// ---- POUs/Tc2 Objects/Signals/Watchdog/FB_SignalWatchdog.TcPOU
FUNCTION_BLOCK FB_SignalWatchdog
VAR_INPUT
	(* Input variables / Eingang Variablen *)
	bEnable					:BOOL;						(* Enable FB signal *)
	bIn						:BOOL;						(* Input signal *)
	tWatchdog				:TIME := t#0s;					(* Watchdog time *)
END_VAR
VAR_OUTPUT
	(* Output variables / Ausgang Variablen *)
	bOut					:BOOL;						(* Output signal *)
	bAlarm					:BOOL;						(* Alarm signal *)
END_VAR
VAR
	(* Enummerations *)

	(* Variables *)


	(* References *)

	(* Interfaces *)

	(* Instances *)
	tofWatchdog				:TOF;

END_VAR

IF NOT bEnable
THEN
	bOut := FALSE;
	bAlarm := FALSE;                       (* Alarm active *)
	
	tofWatchdog(
		IN := tofWatchdog.ET > t#0ms,
	         PT := t#0ms
	);
	
	tofWatchdog(IN := FALSE,
	             PT := t#0ms);

	RETURN;
END_IF;

tofWatchdog(					 (* Dealy input signal *)
	IN := bIn,
	PT := tWatchdog
);

bOut := tofWatchdog.Q;

bAlarm := NOT tofWatchdog.Q;                       (* Set alarm *)

END_FUNCTION_BLOCK

// ---- POUs/Machine/Group_0000 - General/Gr00Control/Gr00Signals/FB_Gr00Signals.TcPOU
FUNCTION_BLOCK FB_Gr00Signals
(*

The function block used to control general signals of the machine.

Constructor: 		Patryk Panylo
Company:		E. Riexinger GmbH
Date:			28.04.2015
Version:			1.00

Date:			Revision:		Who:				Comment
dd.mm.yyyy		x.xx			Initials			comment

*)
VAR_INPUT
	(* Input variables / Eingang Variablen *)
	etMachineMode				:ET_MachineMode;			(* Machine mode *)
	etMachineState				:ET_MachineState;			(* Machine state *)
	bMachineRunning				:BOOL;						(* Machine running / Maschine lauft *)
	stAlarm						:ST_Alarm;					(* Current status of alarms *)
END_VAR
VAR_OUTPUT
	(* Output variables / Ausgang Variablen *)
	bBulbRed					:BOOL;						(* Signal column bulb "stop" or "error" / Signallampe "Stop" oder "Fehler" *)
	bBulbYellow					:BOOL;						(* Signal column bulb "warning" or "message" / Signallampe "Warnung" oder "Message" *)
	bBulbGreen					:BOOL;						(* Signal column bulb "automatic" / Signallampe "Automatik" *)
	bBulbBtnStop					:BOOL;						(* Signal button bulb "stop" / Signallampe "Stop" *)
	bBulbBtnHome				:BOOL;						(* Signal button bulb "home" / Signallampe "Grundstellung" *)
	bBulbBtnStart					:BOOL;						(* Signal button bulb "start" / Signallampe "Start" *)
	bHorn						:BOOL;						(* Signal horn / Signalhupe *)
	stBlinker						:ST_Blinker;
END_VAR
VAR_IN_OUT
	(* Input Output variables / Ausgang Variablen *)

END_VAR
VAR
	(* Enummerations *)

	(* Variables *)
	nIdxHorn						:INT;

	(* References *)

	(* Interfaces *)

	(* Instances *)
	fbBlinker						:FB_Blinker;
	rtHorn						:R_TRIG;
	tonDelay						:TON;

END_VAR
VAR CONSTANT
	nHornRepeat					:INT := 3;
END_VAR


A_Blinker();
A_SignalColumn();
A_SignalButton();
A_Horn();

ACTION A_Blinker:

(* Blinker frequency division *)
fbBlinker(
    stBlinker => stBlinker
);
END_ACTION

ACTION A_Horn:

(* Signal horn / Signalhupe *)
IF stBlinker.Q1
     AND nIdxHorn < nHornRepeat
THEN
	bHorn := (stAlarm.bFatalError OR stAlarm.bError);

ELSIF NOT stBlinker.Q1
THEN
	bHorn := FALSE;
END_IF;

rtHorn(CLK := bHorn);
IF rtHorn.Q
THEN
	nIdxHorn := nIdxHorn + 1;
END_IF;

tonDelay(
	IN := nIdxHorn >= nHornRepeat,
	PT := t#60s
);

IF (tonDelay.Q
    AND nHornRepeat > 0)
    OR NOT (stAlarm.bFatalError OR stAlarm.bError)
THEN
	nIdxHorn := 0;
END_IF;
END_ACTION

ACTION A_SignalButton:

(* Signal button bulb "stop" / Signallampe "Stop" *)
bBulbBtnStop := bBulbRed;

(* Signal button bulb "home" / Signallampe "Grundstellung" *)
bBulbBtnHome := (
	(etMachineMode = ET_MachineMode_eHome
	 AND NOT bMachineRunning)
	OR
	(etMachineMode = ET_MachineMode_eHome
	 AND bMachineRunning
	 AND stBlinker.Q1)
);

(* Signal button bulb "start" / Signallampe "Start" *)
bBulbBtnStart := (
	(etMachineMode = ET_MachineMode_eAutomatic
	 AND bMachineRunning)
	OR
	(etMachineMode = ET_MachineMode_eHome
	 AND bMachineRunning
	 AND NOT stBlinker.Q1)
);
END_ACTION

ACTION A_SignalColumn:

(* Signal column bulb "stop" or "error" / Signallampe "Stop" oder "Fehler" *)
bBulbRed := SEL(
	stAlarm.bFatalError OR stAlarm.bError,
	NOT bMachineRunning,
	stBlinker.Q1
);

(* Signal column bulb "warning" or "message" / Signallampe "Warnung" oder "Message" *)
bBulbYellow := (
	NOT stBlinker.Q1
	AND (stAlarm.bWarning OR stAlarm.bMessage)
);

(* Signal column bulb "automatic" / Signallampe "Automatik" *)
bBulbGreen := (
	(etMachineMode = ET_MachineMode_eAutomatic
	 AND bMachineRunning)
	OR
	(etMachineMode = ET_MachineMode_eHome
	 AND bMachineRunning
	 AND stBlinker.Q1)
);
END_ACTION

END_FUNCTION_BLOCK

// ---- POUs/Tc2 Objects/Signals/Generators/FB_Blinker.TcPOU
FUNCTION_BLOCK FB_Blinker
(*

Frequency division

Constructor: 		Patryk Panylo
Company:		E. Riexinger GmbH
Date:			14.11.2012
Version:			1.00

Date:			Revision:		Who:				Comment
dd.mm.yyyy		x.xx			Initials			comment

*)

VAR_INPUT
	tPeriod				:TIME := T#250MS;				(* Blink period *)
	bReset				:BOOL;						(* Reset *)
END_VAR
VAR_OUTPUT
	stBlinker				:ST_Blinker;
END_VAR
VAR
	byInc				:BYTE;
	rtTriger				:R_TRIG;
	ton1					:TON;
	ton2					:TON;
END_VAR

IF bReset
THEN
	byInc := 0;

	ton1(IN := FALSE);
	ton2(IN := FALSE);

	stBlinker.Q0 := 0;
	stBlinker.Q1 := 0;
	stBlinker.Q2 := 0;
	stBlinker.Q3 := 0;
	stBlinker.Q4 := 0;
	stBlinker.Q5 := 0;
	stBlinker.Q6 := 0;
	stBlinker.Q7 := 0;
	
	RETURN;	
END_IF

ton1(IN := NOT ton2.Q, PT:= tPeriod/2);
ton2(IN := ton1.Q, PT := tPeriod/2);

rtTriger(CLK := ton1.Q);
IF rtTriger.Q THEN
	byInc := byInc + 1;
END_IF;

stBlinker.Q0 := byInc.0;
stBlinker.Q1 := byInc.1;
stBlinker.Q2 := byInc.2;
stBlinker.Q3 := byInc.3;
stBlinker.Q4 := byInc.4;
stBlinker.Q5 := byInc.5;
stBlinker.Q6 := byInc.6;
stBlinker.Q7 := byInc.7;

END_FUNCTION_BLOCK

// ---- POUs/Machine/Group_0000 - General/Gr00Control/Gr00Utility/FB_Gr00Utility.TcPOU
FUNCTION_BLOCK FB_Gr00Utility
(*

The function block used to control general utility of the machine.

Constructor: 		Patryk Panylo
Company:		E. Riexinger GmbH
Date:			28.04.2015
Version:			1.00

Date:			Revision:		Who:				Comment
dd.mm.yyyy		x.xx			Initials			comment

*)
VAR_INPUT
	(* Input variables / Eingang Variablen *)
	bSignalStart					:BOOL;						(* Signal "Start" / Signal "Start" *)
	bSignalStop					:BOOL;						(* Signal "Stop" / Signal "Stop" *)
	bSignalAbort					:BOOL;						(* Signal "Abort" / Signal "Abort" *)
	bSignalHome					:BOOL;						(* Signal "Home" / Signal "Grundstellung" *)
	bSignalReference				:BOOL;						(* Signal "Reference" / Signal "Referenz" *)
	bSignalReset					:BOOL;						(* Signal "Reset" / Signal "Reset *)
	bSignalMachinePurge			:BOOL;						(* Machine purge *)
	bAutoStartRelease			:BOOL;						(* Auto start release *)
	bHomeStartRelease			:BOOL;						(* Home start release *)
	bAutoToHome				:BOOL;						(* If auto completed go to home *)
	bHomeCompleted				:BOOL;						(* Home completed signal *)
	bAutoCompleted				:BOOL;						(* Auto completed signal *)
	bAllDoorsClosed 				:BOOL;						(* All doors closed *)
	bAllDoorsLocked 				:BOOL;						(* All doors locked *)
	bLightCurtainOk				:BOOL;						(* Light curtain ok *)
	bExeCounter					:BOOL;						(* Execute counter *)
	bResetCounterUser			:BOOL;						(* Reset counter user *)
	bStartTime					:BOOL;						(* Start measurement of cylce time *)
	bStopTime					:BOOL;						(* Stop measurement of cylce time *)
	bLifetimeOn					:BOOL;						(* Lifetime on *)
	bResetLifetimeAll				:BOOL; 						(* Reset all counters *)
	sLifetimeFilePath				:STRING;					(* File path for life time *)
	sLifetimeFileName			:STRING;					(* File name for life time *)
	bWritePersistent				:BOOL;						(* Write persistent data *)
	bDownTraceDataExe 			:BOOL;						(* Download traceability data *)
	stTraceability					:ST_Traceability;				(* Traceability data *)
	tAdsTimeOut 					:TIME := t#2s;					(* Timout for ads commands *)
END_VAR
VAR_OUTPUT
	(* Output variables / Ausgang Variablen *)
	etMachineMode				:ET_MachineMode;			(* Machine mode *)
	etMachineState				:ET_MachineState;			(* Machine state *)
	bModeAutomatic				:BOOL;						(* Machine mode automatic *)
	bModeHome					:BOOL;						(* Machine mode home *)
	bModeManual				:BOOL;						(* Machine mode manual *)
	bMachineRunning				:BOOL;						(* Machine running *)
	bMachineStandstill			:BOOL;						(* Machine standstill *)
	bMachinePurge				:BOOL;						(* Machine purge *)
	bConfirmAlarm				:BOOL;						(* Alarm confirm *)
	rActOverride					:REAL;						(* Actual override *)
	lrLifetimeAll					:LREAL;						(* Lifetime *)
	lrLifetimeAfterTrunOn			:LREAL;						(* Time after turn on *)
	lrActCycleTime				:LREAL;						(* Actual cycle time *)
	dwCycleTime					:DWORD;					(* Cycletime in 0.01sec / Zykluszeit in 0.01Sekunden *)
END_VAR
VAR_IN_OUT
	(* Input Output variables / Ausgang Variablen *)
	etMachineModeReq			:ET_MachineMode;			(* Machine mode request *)
	rGlobalOverride				:REAL;						(* Global override *)
	udnCounterTotal				:UDINT;						(* Total counter *)
	udnCounterUser				:UDINT;						(* Total counter *)
END_VAR
VAR
	(* Enummerations *)

	(* Variables *)
	nIRHSCtrlCnt					:INT;
	nIRHSZoneCnt				:INT;
	lrIRHSSetpointLeftSide			:LREAL;
	lrIRHSSetpointRightSide		:LREAL;

	bTraceExe					:BOOL;
	ftTraceExe					:F_TRIG;
	rtDownTraceDataExe			:R_TRIG;
	rtDownTraceDataReset		:R_TRIG;
	udnTraceSampleCnt			:UDINT;
	udnTraceDataCnt				:UDINT;

	(* References *)

	(* Interfaces *)

	(* Instances *)
	fbModeSelector				:FB_ModeSelector;			(* Mode selector *)
	fbOverride					:FB_Override;					(* Override *)
	fbLifetime					:FB_TimeHoursCounter;		(* Machine lifetime *)
	fbCounterTotal				:FB_Counter;					(* Counter total *)
	fbCounterUser				:FB_Counter;					(* Counter user *)
	rtResetCounterUser			:R_TRIG;						(* Reset counter user *)
	fbCylceTime					:FB_Timer;					(* Machine cycle time *)
	fbSUPS						:FB_S_UPS_CX51x0;			(*  The function block FB_S_UPS_CX51x0 can be used on CX devices with one-second UPS to control the one-second UPS from the PLC *)
	fbWritePersistentData			:WritePersistentData;			(*  Write Persistent *)
	fbGetCurTaskIdx				:GETCURTASKINDEX;			(* This function block finds the task index of the task from which it is called *)
	fbRTC						:FB_RTC;					(* Get current time *)
	fbTraceability					:FB_Traceability;				(* Traceability *)
	rtMachinePurge				:R_TRIG;
	SystemTaskInfoArr: INT;
END_VAR


A_OperationMode();
A_Override();
A_Counter();
A_CycleTime();
A_MachinePurge();
A_Persistent();
A_PlcTaskSystemInfo();
A_RTC();
A_Traceability();

ACTION A_Counter:

(* Hours counter *)
fbLifetime(
	bEnable := TRUE,
	bDeleteAll := bResetLifetimeAll,
	sAmsNetId := sgAmsNetId,
	bCount := bLifetimeOn,
	bSave := FALSE,
	sFilePath := sLifetimeFilePath,
	sFileName := sLifetimeFileName,
	tSaveIntervall := t#5m,
	tTimeout := tAdsTimeOut,
	lrAllOverHours => lrLifetimeAll,
	lrNoRetainHours => lrLifetimeAfterTrunOn,
 );

(* General counter *)
fbCounterTotal(
	bEnable := TRUE,
	bExecute := bExeCounter,
	bReset := fbCounterTotal.bOverflow,
	udnCounter := udnCounterTotal
);

rtResetCounterUser(CLK:= bResetCounterUser);

fbCounterUser(
	bEnable := TRUE,
	bExecute := bExeCounter,
	bReset := rtResetCounterUser.Q
			 OR fbCounterUser.bOverflow,
	udnCounter := udnCounterUser
);
END_ACTION

ACTION A_CycleTime:

(* Cylce time *)
fbCylceTime(
	bEnable := TRUE,
	bReset := FALSE,
	bStartStop := bStartTime
			        AND bModeAutomatic,
	bStop := bStopTime
		        OR bMachineStandstill,
	tMaxTime := ,
	stRefTime => ,
	stActTime => ,
	stRestTime =>
);

dwCycleTime := fbCylceTime.stActTime.dwDeciSec;
END_ACTION

ACTION A_MachinePurge:

rtMachinePurge(CLK := 	bSignalMachinePurge);

IF NOT bModeAutomatic
     OR bAutoCompleted
THEN
	bMachinePurge := FALSE;

ELSIF rtMachinePurge.Q
THEN
	bMachinePurge := TRUE;
END_IF
END_ACTION

ACTION A_OperationMode:

(* Operation mode control *)
fbModeSelector(
	bStart := bSignalStart,
	bStop := bSignalStop,
	bAbort := bSignalAbort,
	bHome := bSignalHome,
	bReset := bSignalReset,
	bReference := bSignalReference,
	bAutoStartRelease := bAutoStartRelease,
	bHomeStartRelease := bHomeStartRelease,
	bAutoToHome := bAutoToHome,
	bHomeCompleted := bHomeCompleted,
	bAutoCompleted := bAutoCompleted,
	bAllDoorsClosed  := bAllDoorsClosed,
	bAllDoorsLocked := bAllDoorsLocked,
	bLightCurtainOk := bLightCurtainOk,
	etMachineMode => etMachineMode,
	etMachineState => etMachineState,
	bModeAutomatic => bModeAutomatic,
	bModeHome => bModeHome,
	bModeManual => bModeManual,
	bMachineRunning => bMachineRunning,
	bMachineStandstill => bMachineStandstill,
	bConfirmAlarm => bConfirmAlarm,
	etMachineModeReq := etMachineModeReq
);
END_ACTION

ACTION A_Override:

(* Override control *)
fbOverride(
	bEnable := TRUE,
	bBypassAccDec := bModeManual,
	bSetOverideMax := bModeAutomatic,
	rAcc := rgGr00AdsOverrideAcc,
	rDec := rgGr01AdsOverrideDec,
	rSetOverride := rGlobalOverride,
	rActOverride => rActOverride
);
END_ACTION

ACTION A_Persistent:

(*  The function block FB_S_UPS_CX51x0 can be used on CX devices with one-second UPS to control the one-second UPS from the PLC *)
fbSUPS(
	sNetID := sgAmsNetId,													(* AmsNetID of the controller. *)
	iPLCPort := AMSPORT_R0_PLC_RTS1,									(* Port number of the PLC runtime system (AMSPORT_R0_PLC_RTS1 = 801, AMSPORT_R0_PLC_RTS2 = 811, AMSPORT_R0_PLC_RTS3 = 821, AMSPORT_R0_PLC_RTS4 = 831). *)
	iUPSPort := 16#588,													(* Port number via which the UPS status is read (standard value is 16#588) *)
	tTimeout := DEFAULT_ADS_TIMEOUT,									(* ADS Timeout *)
	eUpsMode := eSUPS_WrPersistData_Shutdown,							(* The eUpsMode defines whether persistent data are to be written and whether a QuickShutdown is to be performed.
																		Standard value is eSUPS_WrPersistData_Shutdown, i.e. with writing of the persistent data and then QuickShutdown. See E_S_UPS_Mode. *)
	ePersistentMode := SPDM_2PASS,										(* Mode for the writing of the persistent data. Standard value is SPDM_2PASS *)
	tRecoverTime := t#10s													(* Time after which the UPS reverts to the PowerOK status in the case of UPS modes without shutdown.
																	   	    The tRecoverTime must be somewhat longer than the maximum holding time of the UPS, since the UPS switches off even when the voltage returns. *)
);


(* If persistent variables are defined in one of the PLC's runtime systems, then their current values are stored in a file in the TwinCAT\Boot directory when the TwinCAT system stops (after the last PLC cycle). *)
fbWritePersistentData(
	NETID := sgAmsNetId,
	PORT := AMSPORT_R0_PLC_RTS1,
	START := bWritePersistent
			   AND NOT fbWritePersistentData.BUSY,
	TMOUT := DEFAULT_ADS_TIMEOUT
);
END_ACTION

ACTION A_PlcTaskSystemInfo:

fbGetCurTaskIdx();

// lrActCycleTime := UDINT_TO_LREAL(SystemTaskInfoArr[fbGetCurTaskIdx.index].cycleTime) / 10000000;




fbGetCurTaskIdx();

GVL._PlcTaskSystemInfo := _TaskInfo[fbGetCurTaskIdx.index];

lrActCycleTime := UDINT_TO_LREAL(_TaskInfo[fbGetCurTaskIdx.index].CycleTime) / 10000000;
END_ACTION

ACTION A_RTC:

fbRTC(
	stDateTime => stgGr00DateTime
);
END_ACTION

ACTION A_Traceability:

stTraceability.sDateTime := stgGr00DateTime.sDateTime;

stTraceability.stSettings.sPath := sTracePath(*CONCAT(CONCAT(sTracePath,fbRTC.sDate),'\')*);
stTraceability.stSettings.sFileName := stgGr00DateTime.sDateTime;
stTraceability.stSettings.sFileExtension := sTraceFileExtension;

rtDownTraceDataReset(
	CLK := bModeAutomatic
);

IF rtDownTraceDataReset.Q
THEN
	udnTraceSampleCnt := 0;
	MEMSET(ADR(stTraceability.arstData), 0, SIZEOF(stTraceability.arstData));
END_IF

rtDownTraceDataExe(
	CLK := bTraceEnable
		    AND bDownTraceDataExe
);

IF rtDownTraceDataExe.Q
     AND udnTraceSampleCnt < udnTraceSampleMax
THEN
	udnTraceDataCnt := 0;
	udnTraceSampleCnt := udnTraceSampleCnt +1;
	(*1*)
	udnTraceDataCnt := udnTraceDataCnt + 1;
	stTraceability.arstData[udnTraceSampleCnt,udnTraceDataCnt].sName := 'Time';
	stTraceability.arstData[udnTraceSampleCnt,udnTraceDataCnt].sValue := stgGr00DateTime.sDateTime;
	stTraceability.arstData[udnTraceSampleCnt,udnTraceDataCnt].sUnit := '';

	(*2*)
	udnTraceDataCnt := udnTraceDataCnt + 1;
	stTraceability.arstData[udnTraceSampleCnt,udnTraceDataCnt].sName := 'Cntr';
	stTraceability.arstData[udnTraceSampleCnt,udnTraceDataCnt].sValue := UDINT_TO_STRING(stgGr00HMI.stPLCTOHMI.udnCounterTotal);
	stTraceability.arstData[udnTraceSampleCnt,udnTraceDataCnt].sUnit := '';

END_IF

(*ftTraceExe(CLK := bgGr00ModeAutomatic);*)
fbTraceability(
	bEnable := bTraceEnable,
	bExecute := bAutoCompleted
			     (*OR
			     (NOT bAutoCompleted
			      AND (bSignalStop OR bSignalAbort)
			      AND ftTraceExe.Q)*)
			     OR bTraceExe,
	stTraceability := stTraceability
);
END_ACTION

END_FUNCTION_BLOCK

// ---- POUs/Tc2 Objects/Automation/OperationMode/FB_ModeSelector.TcPOU
FUNCTION_BLOCK FB_ModeSelector
(*

The function block used to control opration mode.

Constructor: 		Patryk Panylo
Company:		E. Riexinger GmbH
Date:			23.04.2015
Version:			1.00

Date:			Revision:		Who:				Comment
dd.mm.yyyy		x.xx			Initials			comment

*)
VAR_INPUT
	(* Input variables / Eingang Variablen *)
	bStart					:BOOL;						(* Signal start *)
	bStop					:BOOL;						(* Signal stop *)
	bAbort					:BOOL;						(* Signal abort *)
	bHome					:BOOL;						(* Signal home *)
	bReference				:BOOL;						(* Signal reference *)
	bReset					:BOOL;						(* Signal reset *)
	bAutoStartRelease		:BOOL;						(* Auto start release *)
	bHomeStartRelease		:BOOL;						(* Home start release *)
	bAutoToHome			:BOOL;						(* If auto completed go to home *)
	bHomeCompleted			:BOOL;						(* Home completed *)
	bAutoCompleted			:BOOL;						(* Auto completed *)
	bAllDoorsClosed 			:BOOL;						(* All doors closed *)
	bAllDoorsLocked 			:BOOL;						(* All doors locked *)
	bLightCurtainOk			:BOOL;						(* Light curtain ok *)
END_VAR
VAR_OUTPUT
	(* Output variables / Ausgang Variablen *)
	etMachineMode			:ET_MachineMode;			(* Machine mode enum variable *)
	etMachineState			:ET_MachineState;			(* Machine state enum variable *)
	bModeAutomatic			:BOOL;						(* Machine mode automatic *)
	bModeHome				:BOOL;						(* Machine mode home *)
	bModeManual			:BOOL;						(* Machine mode manual *)
	bMachineRunning			:BOOL;						(* Machine running *)
	bMachineStandstill		:BOOL;						(* Machine standstill *)
	bConfirmAlarm			:BOOL;						(* Confirm alarm *)
END_VAR
VAR_IN_OUT
	etMachineModeReq		:ET_MachineMode;			(* Machine mode request enum variable *)
END_VAR
VAR
	(* Enummerations *)

	(* Variables *)
	etMachinePrvState		:ET_MachineState;			(* Machine previous active state enum variable *)
	bModeExecute			:BOOL;						(* Mode execute *)
	bSafetyCompleted		:BOOL;						(* Safety completed *)

	(* References *)

	(* Interfaces *)

	(* Instances *)
	rtStart					:R_TRIG;
	rtStop					:R_TRIG;
	rtAbort					:R_TRIG;
END_VAR


bConfirmAlarm := bReset;
bSafetyCompleted := bAllDoorsLocked				(* Safety completed *)
				      AND bLightCurtainOk;

IF bHome
THEN
	etMachineModeReq := ET_MachineMode_eHome;

END_IF;

IF bHomeCompleted
THEN
	IF etMachineMode = ET_MachineMode_eHome                          	 (* Set auto mode *)
	    AND etMachinePrvState <> ET_MachineState_eAutoExe
	    AND etMachinePrvState <> ET_MachineState_eAutoSteppingExe
	    AND etMachinePrvState <> ET_MachineState_eAutoSteppingNoExe
	    AND bModeExecute
	THEN
		etMachineModeReq := ET_MachineMode_eAutomatic;

	END_IF;
ELSE
	IF etMachineModeReq <> ET_MachineMode_eManual                   	 (* Set home mode *)
	THEN
		etMachineModeReq := ET_MachineMode_eHome;
	
	END_IF;
END_IF;

IF (etMachineModeReq <> etMachineMode)                                    		(* Stop always if changed mode *)
THEN
	(*bStart := FALSE *)
	bStop := TRUE;

	IF (etMachineMode = ET_MachineMode_eAutomatic
	      AND etMachineModeReq = ET_MachineMode_eStepping)
	     OR
	     (etMachineMode = ET_MachineMode_eStepping
	      AND etMachineModeReq = ET_MachineMode_eAutomatic)
	THEN
		bStop := FALSE;
	END_IF;

	etMachineMode := etMachineModeReq;
END_IF;

rtStart(CLK := bStart);								(* Check start *)

rtStop(CLK := bStop								(* Check stop *)
		        OR bAbort
		        OR bAutoCompleted
		        OR (NOT bSafetyCompleted AND bMachineRunning));
rtAbort(CLK := bAbort);

IF rtStop.Q
THEN
	bModeExecute := FALSE;

	IF bAutoToHome
	     AND bAutoCompleted
	     OR(bMachineRunning
		    AND bModeAutomatic
		    AND bHomeCompleted
		    AND NOT bAutoCompleted)
	THEN
		etMachineModeReq := ET_MachineMode_eHome;
	END_IF

ELSIF rtStart.Q
	    AND bAllDoorsClosed
	    AND bLightCurtainOk
	    AND NOT bStop
	    AND NOT bAbort
	    AND ((etMachineMode = ET_MachineMode_eHome AND SEL(
															etMachineState = ET_MachineState_eHomeExe
															OR etMachineState = ET_MachineState_eHomeRefExe,
															bHomeStartRelease, TRUE))
	    	       OR ((etMachineMode = ET_MachineMode_eAutomatic
			        OR etMachineMode = ET_MachineMode_eStepping) AND SEL(
																		etMachineState = ET_MachineState_eAutoExe
																		OR etMachineState = ET_MachineState_eAutoSteppingExe
																		OR etMachineState = ET_MachineState_eAutoSteppingNoExe,
															bAutoStartRelease, TRUE)))
THEN
	bModeExecute := TRUE;

END_IF;

bStart := FALSE;
bStop := FALSE;

CASE etMachineMode
OF
	ET_MachineMode_eAutomatic:            (* Statement section automatic *)
		bModeAutomatic := TRUE;
		bModeHome := FALSE;
		bModeManual := FALSE;

		IF bModeExecute
		     AND bSafetyCompleted
		THEN
			etMachineState := ET_MachineState_eAutoExe;
			etMachinePrvState := etMachineState;
		ELSE
		 	etMachineState := ET_MachineState_eIdle;
		END_IF;
	    
	ET_MachineMode_eStepping:             (* Statement section stepping *)
		bModeAutomatic := TRUE;
		bModeHome := FALSE;
		bModeManual := FALSE;

		IF bModeExecute
		     AND bSafetyCompleted
		THEN
			IF rtStart.Q
			THEN
				etMachineState := ET_MachineState_eAutoSteppingExe;
			ELSE
				etMachineState := ET_MachineState_eAutoSteppingNoExe;
			END_IF;

			etMachinePrvState := etMachineState;
		ELSE
			etMachineState := ET_MachineState_eIdle;
		END_IF;

	ET_MachineMode_eHome:                 (* Statement section home  *)
		bModeAutomatic := FALSE;
		bModeHome := TRUE;
		bModeManual := FALSE;

		IF bModeExecute
		     AND bSafetyCompleted
		THEN
			IF bReference
			THEN
				etMachineState := ET_MachineState_eHomeRefExe;
			ELSE
				etMachineState := ET_MachineState_eHomeExe;
			END_IF;

			etMachinePrvState := etMachineState;
		ELSE
			etMachineState := ET_MachineState_eIdle;
		END_IF;

	ET_MachineMode_eManual:              (* Statement section manual  *)
		bModeExecute := FALSE;
		bModeAutomatic := FALSE;
		bModeHome := FALSE;
		bModeManual := TRUE;

		etMachineState := ET_MachineState_eIdle;

	ELSE
		bModeExecute := FALSE;
		bModeAutomatic := FALSE;
		bModeHome := FALSE;
		bModeManual := FALSE;
	    
	    	etMachineState := ET_MachineState_eUndefined;
        
END_CASE;

bMachineRunning := bModeExecute
		                       AND etMachineMode <> ET_MachineMode_eManual
		                       AND etMachineMode <> ET_MachineMode_eIdle
		                       AND etMachineMode <> ET_MachineMode_eUndefined;
                    
bMachineStandstill := NOT bMachineRunning;

END_FUNCTION_BLOCK

// ---- POUs/Tc2 Objects/Automation/Axis/Override/FB_Override.TcPOU
FUNCTION_BLOCK FB_Override
(*

The function block used to control override of axis.

Constructor: 		Patryk Panylo
Company:		E. Riexinger GmbH
Date:			23.04.2015
Version:			1.00

Date:			Revision:		Who:				Comment
dd.mm.yyyy		x.xx			Initials			comment

*)
VAR_INPUT
	(* Input variables / Eingang Variablen *)
	bEnable						:BOOL;						(* Signal FB enable *)
	bBypassAccDec				:BOOL;						(* Bypassing acceleratin und deceleration rActOverride = rSetOverride *)
	bSetOverideMax				:BOOL;						(* Set maximum override *)
	rAcc							:REAL;						(* Accerlation of Override [%/s] *)
	rDec						:REAL;						(* Decerlation of Override [%/s] *)
END_VAR
VAR_OUTPUT
	(* Output variables / Ausgang Variablen *)
	rActOverride					:REAL;						(* Actual Override *)
END_VAR
VAR_IN_OUT
	rSetOverride					:REAL;						(* Set Override *)
END_VAR
VAR
	(* Enummerations *)

	(* Variables *)
	rSetOverrideInternal			:REAL;						(* Internal Set Override limited *)
	rAccOverridePerCycle			:REAL;						(* Override accerleration per cycle *)
	rDecOverridePerCycle			:REAL;						(* Override deceleration per cycle *)
	tCycleTime					:TIME;						(* Detected cycle Time *)
	bFirstTime					:BOOL;						(* First run *)

	(* References *)

	(* Interfaces *)

	(* Instances *)
	tonChkCycleTime				:TON;						(* Check cycle time *)
	rtSetOverideMax				:R_TRIG;
END_VAR
VAR CONSTANT
	rMIN_OVERRIDE				:REAL := 0.0;					(* Minimum override *)
	rMAX_OVERRIDE				:REAL := 100.0;				(* Maximum override *)
	rACC_MIN					:REAL := 0.1;					(* Minimum accerleration *)
	rDEC_MIN					:REAL := 0.1;					(* Minimum decerleration *)
	tMAX_CYCLE_TIME			:TIME := t#1s;					(* Maximum cycle time *)
END_VAR

IF NOT bEnable
THEN
	bFirstTime := FALSE;								(* First run *)
	rActOverride := 100.0;								(* Set Override *)
	RETURN;
END_IF;

IF NOT bFirstTime                                             					 (* First run after bEnable *)
THEN
	tonChkCycleTime(					   				 (* Start Timer to check  cycle time *)
		IN := TRUE,
		PT := tMAX_CYCLE_TIME
	);
	
	IF tonChkCycleTime.ET <> t#0s                              			 (* Timer was running one circle *)
	THEN
		tCycleTime := tonChkCycleTime.ET;                     		 (* Detectet circle time *)

		tonChkCycleTime(					 			 (* Stop Timer *)
			IN := FALSE,
			PT := tMAX_CYCLE_TIME
		);

		bFirstTime := TRUE;                                     			(* First run *)
	END_IF;
END_IF;

(* Set max overide *)
rtSetOverideMax(CLK := bSetOverideMax);
IF rtSetOverideMax.Q
THEN
	rSetOverride := rMAX_OVERRIDE;
END_IF

(* Check Limits *)
rSetOverrideInternal := LIMIT(                      					 (* Internal Override Limited *)
	rMIN_OVERRIDE,              							 (* Minimum Override *)
	rSetOverride,              							 	 (* Set Override *)
	rMAX_OVERRIDE               							 (* Maximum Overide *)
);

IF bBypassAccDec
THEN
	rActOverride := rSetOverrideInternal;                  			 (* Actual Override = Set Override *)
ELSE
	IF tCycleTime <> t#0s
	THEN

		A_Acceleration();

		A_Deceleration();

	END_IF;
END_IF;

ACTION A_Acceleration:

IF rSetOverrideInternal > rActOverride                          	(* Override has to be added *)
THEN
	(* Check if accerlaeration zero *)
	IF rAcc <= 0
	THEN
		rAcc := rACC_MIN;                                         	(* Set accerlaeration to minimum *)
	END_IF;

	(* Calculate Accerleration per cycle *)
	rAccOverridePerCycle := rAcc / (TIME_TO_REAL(tMAX_CYCLE_TIME)
							     / TIME_TO_REAL(tCycleTime));
	
	rActOverride := rActOverride + rAccOverridePerCycle;        (* Add Override *)
	IF rActOverride > rSetOverrideInternal                      		 (* Actoverride  run over Set Override ? *)
	THEN
		rActOverride := rSetOverrideInternal;             (* Set  Override equal *)
	END_IF;
END_IF;
END_ACTION

ACTION A_Deceleration:

IF rSetOverrideInternal < rActOverride                             (* Override has to subed *)
THEN
	(* Check if decerlaeration zero *)
	IF rDec <= 0
	THEN
		rDec := rDEC_MIN;                                         	(* Set decerlaeration to minimum *)
	END_IF;

	(* Calculate decerleration per cycle *)
	rDecOverridePerCycle := rDec / (TIME_TO_REAL(tMAX_CYCLE_TIME) /
								TIME_TO_REAL(tCycleTime));
	
	rActOverride := rActOverride - rDecOverridePerCycle;        (* Sub Override *)
	IF rActOverride < rSetOverrideInternal                        		 (* Actoverride  run over Set Override ? *)
	THEN
	    rActOverride := rSetOverrideInternal;                  (* Set  Override equal *)
	END_IF;
END_IF;
END_ACTION

END_FUNCTION_BLOCK

// ---- POUs/Tc2 Objects/Measurements/Counter/FB_TimeHoursCounter.TcPOU
FUNCTION_BLOCK FB_TimeHoursCounter
(*

Function block to read and write elapsed time in/from file.
If sFileName or sFilePath  or sFileSuffix is empty then save function is diabled and generate error.

Constructor: 		Patryk Panylo
Company:		E. Riexinger GmbH
Date:			17.03.2014
Version:			1.00

Date:			Revision:		Who:				Comment
dd.mm.yyyy		x.xx			Initials			comment

*)

VAR_INPUT
	(* Variables *)
	bEnable							:BOOL;							(* Enable FB *)
	sAmsNetId 						:STRING := ''; 						(* Ams Net ID of file to read/write *)
	bCount							:BOOL; 							(* If true then count time else save current time *)
	bSave							:BOOL;							(* Save current hours counter *)
	bReset							:BOOL; 							(* Reset counter *)
	bDeleteAll						:BOOL; 							(* Delete all counters since beginning *)
	sFilePath						:STRING := 'C:\TwinCAT\Plc\';		(* File path *)
	sFileName						:STRING := 'default';				(* File name *)
	tSaveIntervall						:TIME := t#3m;						(* Intervall to save counter hours. If equal 0 then intervall is off *)
	tTimeout							:TIME := t#3s;						(* ADS timeout *)
END_VAR
VAR_OUTPUT
	(* Variables *)
	lrAllOverHours					:LREAL; 							(* All over counter hours *)
	lrAfterResetHours					:LREAL; 							(* Counter hours since last reset *)
	lrNoRetainHours					:LREAL; 							(* No retain counter hours *)
	bError							:BOOL;							(* Program error *)
	udnErrNo						:UDINT;							(* Error number *)
END_VAR
VAR
	(* Enummerations *)
	etRWStep						:(eReadHours, eChkRead, eWFWrite, eWriteHours, eChkWrite, eError );

	(* Variables *)
	bFirstTime						:BOOL;
	arlrCycleTimeAsHour				:ARRAY[0..2] OF LREAL;			(* Current cycle time as hours *)
	stRetainHours					:ST_TimeHoursCounter;

	(* Instances *)
	ftCount							:F_TRIG;
	rtSave							:R_TRIG;
	rtReset							:R_TRIG;
	rtDeleteAll						:R_TRIG;

	fbFileHandler						:FB_FileHandlerBinary;				(* File handler *)
	fbGetSystemTime					:GETSYSTEMTIME;				(* Detects System time *)
	tonWriteIntervall					:TON;							(* Timer for Save intervall control *)

END_VAR

IF NOT bEnable				(* Enable FB *)
THEN
	fbFileHandler(
		bEnable := FALSE,
		bExecute := FALSE,
		bFileRead := FALSE,
		bFileWrite := FALSE
	);

	bFirstTime := FALSE;
	bError := FALSE;			(* Program error *)
	udnErrNo := 0;				(* Error number *)

	RETURN;
END_IF


IF NOT bFirstTime
THEN
	(* Produce the file directory name *)
	fbFileHandler.sFilePath := sFilePath;
	fbFileHandler.sFileName := sFileName;
	fbFileHandler.sFileSuffix := 'thc';

	(* Get cycle time as hours *)
	A_GetCycleTime();

	tonWriteIntervall(
		IN := FALSE,
		PT:= tSaveIntervall
	);

	etRWStep := eReadHours;

	RETURN;
END_IF


(* Read / Write all over hours *)
CASE etRWStep OF

	eReadHours:
		fbFileHandler.bExecute := TRUE;
		fbFileHandler.bFileRead := TRUE;
		fbFileHandler.bFileWrite := FALSE;

		IF fbFileHandler.bBusy
		THEN
			etRWStep := eChkRead;

		END_IF

	eChkRead:
		IF NOT fbFileHandler.bBusy
		THEN
			IF  fbFileHandler.bError
			THEN
				fbFileHandler.bExecute := FALSE;
				fbFileHandler.bFileRead := FALSE;
				fbFileHandler.bFileWrite := FALSE;

				etRWStep := eWFWrite;				(* Next step *)

			ELSE
				fbFileHandler.bExecute := FALSE;
				fbFileHandler.bFileRead := FALSE;
				fbFileHandler.bFileWrite := FALSE;

				etRWStep := eWFWrite;				(* Next step *)

			END_IF
		END_IF

	eWFWrite:
		ftCount(
			CLK :=  bCount AND NOT bReset AND NOT bDeleteAll
		);

		rtSave(
			CLK := bSave AND NOT bReset AND NOT bDeleteAll
		);


		tonWriteIntervall(IN := tSaveIntervall > t#0s);

		IF ftCount.Q
		     OR rtSave.Q
		     OR tonWriteIntervall.Q
		THEN
			tonWriteIntervall(IN := FALSE);

			etRWStep := eWriteHours;								(* Next step *)

		END_IF

	eWriteHours:
		fbFileHandler.bExecute := TRUE;
		fbFileHandler.bFileRead := FALSE;
		fbFileHandler.bFileWrite := TRUE;

		IF fbFileHandler.bBusy
		THEN
			etRWStep := eChkWrite;								(* Next step *)

		END_IF

	eChkWrite:
		IF NOT fbFileHandler.bBusy
		THEN
			IF  fbFileHandler.bError
			THEN
				etRWStep := eError;								(* Next step *)

			ELSE
				fbFileHandler.bExecute := FALSE;
				fbFileHandler.bFileRead := FALSE;
				fbFileHandler.bFileWrite := FALSE;

				etRWStep := eWFWrite;							(* Next step *)

			END_IF
		END_IF

	eError:
		fbFileHandler.bExecute := FALSE;
		fbFileHandler.bFileRead := FALSE;
		fbFileHandler.bFileWrite := FALSE;

END_CASE


(* Counting hours *)
IF bCount
    AND NOT fbFileHandler.bFileRead
THEN
	stRetainHours.lrAllOverHours := stRetainHours.lrAllOverHours + arlrCycleTimeAsHour[0];
	stRetainHours.lrAfterResetHours := stRetainHours.lrAfterResetHours + arlrCycleTimeAsHour[0];
	lrNoRetainHours := lrNoRetainHours + arlrCycleTimeAsHour[0];
END_IF


(* Write / read  file *)
fbFileHandler(
	bEnable := TRUE,
	dwDataBuffer := ADR(stRetainHours),
	udnDataBufLen := SIZEOF(stRetainHours),
	tTimeout := tTimeout,
	bError => bError,
	udnErrNo => udnErrNo
);

rtReset(
	CLK := NOT bSave AND bReset
);
IF rtReset.Q
THEN
	stRetainHours.lrAfterResetHours := 0;
	lrNoRetainHours := 0;
END_IF

rtDeleteAll(
	CLK := NOT bSave AND bDeleteAll
);
IF rtDeleteAll.Q
THEN
	stRetainHours.lrAllOverHours := 0;
	stRetainHours.lrAfterResetHours := 0;
	lrNoRetainHours := 0;
END_IF

(* Counter hours mapping *)
lrAllOverHours := stRetainHours.lrAllOverHours;
lrAfterResetHours := stRetainHours.lrAfterResetHours;

ACTION A_GetCycleTime:

(* Calculate system time *)
fbGetSystemTime;
arlrCycleTimeAsHour[0] := UINT64_TO_LREAL(IN := ULARGE_INTEGER(dwHighPart := fbGetSystemTime.timeHiDW, dwLowPart := fbGetSystemTime.timeLoDW))
									/ 10				(* Calculate into mycro seconds *)
									/ 1000			(* Calculate into millis econds *)
									/ 1000			(* Calculate into seconds *)
									/ 60				(* Calculate into minutes *)
									/ 60;				(* Calculate into hours *)


arlrCycleTimeAsHour[2] := arlrCycleTimeAsHour[1];
arlrCycleTimeAsHour[1] := arlrCycleTimeAsHour[0];

IF arlrCycleTimeAsHour[2] > 0
THEN
	arlrCycleTimeAsHour[0] := ABS(arlrCycleTimeAsHour[2] - arlrCycleTimeAsHour[1]);
	arlrCycleTimeAsHour[1] := 0;
	arlrCycleTimeAsHour[2] := 0;

	bFirstTime := TRUE;
END_IF
END_ACTION

END_FUNCTION_BLOCK

// ---- POUs/Tc2 Objects/File/FB_FileHandlerBinary.TcPOU
FUNCTION_BLOCK FB_FileHandlerBinary
(*

This function block is used to read and write binary datas in/from file.

Constructor: 		Patryk Panylo
Company:		E. Riexinger GmbH
Date:			10.06.2013
Version:			1.00

Date:			Revision:		Who:				Comment
dd.mm.yyyy		x.xx			Initials			comment

*)

VAR_INPUT
	bEnable						:BOOL;					(* Enable FB *)
	bExecute					:BOOL;					(* Execute operation *)
	sFilePath					:STRING;				(* File path *)
	sFileName					:STRING;				(* File name *)
	sFileSuffix					:STRING := 'dat';			(* Suffix of file *)
	bFileWrite					:BOOL;					(* Write file *)
	bFileRead					:BOOL;					(* Read file *)
	dwDataBuffer				:PVOID;				(* Contains the address of the buffer containing the data to be read/written ADR *)
	udnDataBufLen				:UDINT;					(* Contains the number of bytes to be written SIZEOF *)
	tTimeout						:TIME := t#1s;				(* States the time before the function is cancelled *)
END_VAR
VAR_OUTPUT
	bBusy						:BOOL;					(* Program busy *)
	bDone						:BOOL;					(* Program done *)
	bError						:BOOL;					(* Program error *)
	udnErrNo					:UDINT;					(* Error number *)
END_VAR
VAR_IN_OUT

END_VAR
VAR
	(* Enummerations *)
	enStep						: (eWaitExecute := 0, eChkFileName,  eChkBufLen, eFileOpen, eChkFileOpen, eFileWrite, eChkFileWrite, eFileRead, eChkFileRead, eFileClose, eChkFileClose, eDone, eError, eNotExecute);			(* Sequence state for open, read/write and close the file *)

	(* Variables *)
	bFirstTime					:BOOL;					(* First PLC cycle *)

	dwMode						:DWORD;				(* Contains the mode in which the file is to be opened *)
	sPathName					:STRING;				(* Contains the path and filename for the file to be opened *)
	hFileHandle					:UINT;					(* File handle *)

	unWriteCounter				:UINT;
	unReadCounter				:UINT;

	(* Instances *)
	fbFileOpen					:FB_FileOpen;			(* File open *)
	fbFileClose					:FB_FileClose;			(* File close *)
	fbFileRead					:FB_FileRead;			(* File read *)
	fbFileWrite					:FB_FileWrite;				(* File write *)

END_VAR

IF NOT bEnable				(* Enable FB *)
THEN
	bFirstTime := FALSE;		(* First PLC cycle *)
	bBusy := FALSE;			(* Program busy *)
	bDone := FALSE;			(* Program done *)
	bError := FALSE;			(* Program error *)
	udnErrNo := 0;				(* Error number *)
	RETURN;
END_IF

IF NOT bFirstTime
THEN
	enStep := eWaitExecute;

	bFirstTime := TRUE;
END_IF


(* Sequence state for open, read/write and close the file *)
CASE enStep
OF

	eWaitExecute:
		IF bExecute
		THEN
			fbFileOpen.bExecute := FALSE;			(* File open *)
			fbFileClose.bExecute := FALSE;			(* File close *)
			fbFileRead.bExecute := FALSE;			(* File read *)
			fbFileWrite.bExecute := FALSE;			(* File write *)

			bDone := FALSE;
			bError := FALSE;
			udnErrNo := 0;

			IF bFileWrite
			THEN
				dwMode := FOPEN_MODEWRITE OR FOPEN_MODEBINARY;

				enStep := eChkFileName;			(* Next step *)

			ELSIF bFileRead
			THEN
				dwMode := FOPEN_MODEREAD OR FOPEN_MODEBINARY;

				enStep := eChkFileName;			(* Next step *)

			ELSE
				RETURN;
			END_IF

			bBusy := TRUE;

		END_IF

	(* Check file name and path *)
	eChkFileName:

		sPathName := CONCAT(
						sFilePath, CONCAT(
									sFileName, CONCAT(
												'.', sFileSuffix)));

		IF sFilePath <> ''
		     AND sFileName <> ''
		     AND sFileSuffix <> ''
		THEN
			enStep := eChkBufLen;			(* Next step *)

		ELSE
			udnErrNo := eChkFileName;

			enStep := eError;				(* Next step *)

		END_IF


	(* Check buffer lenght *)
	eChkBufLen:
		IF udnDataBufLen = 0
		THEN
			enStep := eDone;				(* Next step *)
	
		ELSE
			enStep := eFileOpen;			(* Next step *)
		
		END_IF

	(* Open the file *)
	eFileOpen:
		fbFileOpen.bExecute := TRUE;

		enStep := eChkFileOpen;				(* Next step *)

	(* Check open the file *)
	eChkFileOpen:
		IF NOT fbFileOpen.bBusy
		THEN
			IF NOT fbFileOpen.bError
			THEN
				fbFileOpen.bExecute := FALSE;
				hFileHandle := fbFileOpen.hFile;

				(* Choose write or read datas *)
				IF fbFileOpen.nMode = (FOPEN_MODEWRITE OR FOPEN_MODEBINARY)
				THEN
					enStep := eFileWrite;			(* Next step *)
	
				ELSIF fbFileOpen.nMode = (FOPEN_MODEREAD OR FOPEN_MODEBINARY)
				THEN
					enStep := eFileRead;			(* Next step *)

				ELSE
					enStep := eFileClose;			(* Next step *)
	
				END_IF

			ELSE
				fbFileOpen.bExecute := FALSE;
				udnErrNo := fbFileOpen.nErrId;
	
				enStep := eError;					(* Next step *)
				
			END_IF
		END_IF

	(* Write the file *)
	eFileWrite:
		fbFileWrite.bExecute := TRUE;

		enStep := eChkFileWrite;				(* Next step *)

	(* Check write the file *)
	eChkFileWrite:
		IF NOT fbFileWrite.bBusy
		THEN
			IF (fbFileWrite.cbWrite >= SIZEOF(dwDataBuffer))
			    AND NOT fbFileWrite.bError
			THEN
				fbFileWrite.bExecute := FALSE;
				unWriteCounter := unWriteCounter + 1;

				enStep := eFileClose;				(* Next step *)

			ELSIF  fbFileWrite.bError
			THEN
				fbFileWrite.bExecute := FALSE;
				udnErrNo := fbFileWrite.nErrId;

				enStep := eError;					(* Next step *)
				
			END_IF
		END_IF

	(* Read the file *)
	eFileRead:
		fbFileRead.bExecute := TRUE;

		enStep := eChkFileRead;				(* Next step *)

	(* Check read the file *)
	eChkFileRead:
		IF NOT fbFileRead.bBusy
		THEN
			IF (fbFileRead.cbRead >= SIZEOF(dwDataBuffer))
			     AND NOT fbFileRead.bError
			THEN
				fbFileRead.bExecute := FALSE;
				unReadCounter := unReadCounter + 1;
	
				enStep := eFileClose;				(* Next step *)

			ELSIF  fbFileRead.bError
			THEN
				fbFileRead.bExecute := FALSE;
				udnErrNo := fbFileRead.nErrId;
	
				enStep := eError;					(* Next step *)
				
			END_IF
		END_IF

	(* Close the file *)
	eFileClose:
		fbFileClose.bExecute := TRUE;

		enStep := eChkFileClose;				(* Next step *)

	(* Check close the file *)
	eChkFileClose:
		IF NOT fbFileClose.bBusy
		THEN
			IF NOT fbFileClose.bError
			THEN
				fbFileClose.bExecute := FALSE;
				enStep := eDone;					(* Next step *)

				IF bError
				THEN
					enStep := eError;				(* Next step *)
				END_IF

			ELSE
				fbFileClose.bExecute := FALSE;
				udnErrNo := fbFileClose.nErrId;
	
				enStep := eError;					(* Next step *)
				
			END_IF
		END_IF

	eDone:
		bBusy := FALSE;
		bDone := TRUE;
		bError := FALSE;
		udnErrNo := 0;

		enStep := eNotExecute;					(* Next step *)

	eError:
		IF NOT bError
		     AND hFileHandle <> 0
		THEN
			bDone := FALSE;
			bError := TRUE;

			enStep := eFileClose;					(* Next step *)

		ELSE
			bBusy := FALSE;
			bDone := FALSE;
			bError := TRUE;
	
			enStep := eNotExecute;					(* Next step *)
		END_IF

	eNotExecute:
		IF NOT bExecute
		THEN
			bBusy := FALSE;
			bDone := FALSE;
			bError := FALSE;
			udnErrNo := 0;

			enStep := eWaitExecute;			(* Next step *)

		END_IF

END_CASE


fbFileOpen(
	sNetId := '',
	sPathName := sPathName,
	nMode := dwMode,
	ePath := PATH_GENERIC,
	tTimeout := tTimeout);
fbFileClose(
	sNetId := '',
	hFile := hFileHandle,
	tTimeout := tTimeout );
fbFileWrite(
	sNetId := '',
	hFile := hFileHandle,
	pWriteBuff := dwDataBuffer,
	cbWriteLen := udnDataBufLen,
	tTimeout := tTimeout);
fbFileRead(
	sNetId := '',
	hFile := hFileHandle,
	pReadBuff := dwDataBuffer,
	cbReadLen := udnDataBufLen,
	tTimeout := tTimeout);

END_FUNCTION_BLOCK

// ---- POUs/Tc2 Objects/Measurements/Counter/FB_Counter.TcPOU
FUNCTION_BLOCK FB_Counter
VAR_INPUT
	(* Input variables / Eingang Variablen *)
	bEnable					:BOOL;						(* Enable FB signal *)
	bExecute				:BOOL;						(* Execute signal *)
	bReset					:BOOL;						(* Reset counter *)
END_VAR
VAR_OUTPUT
	(* Output variables / Ausgang Variablen *)
	bOverflow				:BOOL;						(* Overflow *)
	bAlarm					:BOOL;						(* Alarm signal *)
END_VAR
VAR_IN_OUT
	udnCounter				:UDINT;						(* Counter *)
END_VAR
VAR
	(* Enummerations *)

	(* Variables *)


	(* References *)

	(* Interfaces *)

	(* Instances *)
	rtCount					:R_TRIG;
	rtReset					:R_TRIG;

END_VAR

IF NOT bEnable
THEN

    RETURN;
END_IF;

rtReset(CLK := bReset);                    (* Reset rising edge *)

IF rtReset.Q                               		(* Count reset came *)
THEN
	udnCounter := 0;
END_IF;


rtCount(CLK := bExecute);                   		 (* Trigger rising edge *)

IF rtCount.Q                              		  		 (* Count trigger came *)
THEN
	IF udnCounter = 16#FFFFFFFF		 (* Detect counter overflow *)
	THEN
	    	bOverflow := TRUE;                  	 (* Counter overflow *)
	ELSE
	   	 bOverflow := FALSE;              	   	 (* Not counter overflow *)
	END_IF;
	
	udnCounter := udnCounter + 1;            	 (* Increment counter *)
END_IF;

END_FUNCTION_BLOCK

// ---- POUs/Tc2 Objects/Measurements/FB_Timer.TcPOU
FUNCTION_BLOCK FB_Timer
VAR_INPUT
	(* Input variables / Eingang Variablen *)
	bEnable					:BOOL;						(* Enable FB signal *)
	bReset					:BOOL;						(* Reset timer *)
	bStartStop				:BOOL;						(* Timer start stop *)
	bStop					:BOOL;						(* Timer stop *)
	tMaxTime				:TIME := t#1092m;				(* Maximum time *)
END_VAR
VAR_OUTPUT
	(* Output variables / Ausgang Variablen *)
	stRefTime				:ST_Time;						(* Reference time *)
	stActTime				:ST_Time;						(* Actuel time *)
	stRestTime				:ST_Time;						(* Rest time *)
END_VAR
VAR_IN_OUT

END_VAR
VAR
	(* Enummerations *)

	(* Variables *)
	stTime					:ST_Time;						(* Actuel time *)
	bTimeStarted				:BOOL;							(* Meassuare time started *)

	bFirstTime				:BOOL;

	(* References *)

	(* Interfaces *)

	(* Instances *)
	rtReset					:R_TRIG;
	rtStartStop				:R_TRIG;
	rtStop					:R_TRIG;

	tonMeassureTime			:TON;

END_VAR

IF NOT bEnable
THEN
	bTimeStarted := FALSE;
	rtStartStop(CLK := FALSE);
	tonMeassureTime(
		IN := FALSE,                   (* Reset timer *)
		PT := tMaxTime
	);

	bFirstTime := FALSE;
	RETURN;
END_IF;

IF NOT bFirstTime
THEN
	MEMSET(ADR(stActTime), 0, SIZEOF(stActTime));
	MEMSET(ADR(stRestTime), 0, SIZEOF(stRestTime));
	MEMSET(ADR(stTime), 0, SIZEOF(stTime));
	bFirstTime := TRUE;
END_IF;

IF bReset
THEN
	bTimeStarted := FALSE;
	tonMeassureTime(
		IN := FALSE,
	         PT := tMaxTime
	);
    
	MEMSET(ADR(stActTime), 0, SIZEOF(stActTime));
	MEMSET(ADR(stRestTime), 0, SIZEOF(stRestTime));
	MEMSET(ADR(stTime), 0, SIZEOF(stTime));
END_IF;


(* Rising edge start / stop *)
rtStartStop(CLK := bStartStop);

IF rtStartStop.Q                                   				 (* Startsignal trigger *)
THEN
	IF bTimeStarted                              			 (* Meassuare time started *)
	THEN
		bTimeStarted := TRUE;                      	 (* Time measure started *)
		tonMeassureTime(				 (* Stop (reset) timer *)
			IN := FALSE,
		         PT := tMaxTime
		);
		MEMSET(ADR(stTime), 0, SIZEOF(stTime));
	ELSE
		bTimeStarted := TRUE;                    	 (* Time measure started *)
		MEMSET(ADR(stTime), 0, SIZEOF(stTime));
	END_IF;
END_IF;

(* Rising edge stop*)
rtStop(CLK := bStop);

IF rtStop.Q                                        				 (* Stop timer *)
THEN
	bTimeStarted := FALSE;                        	 	 (* Time measure stoped *)
END_IF;

(* Start timer *)
tonMeassureTime(
	IN := bTimeStarted,
	PT := tMaxTime
);

(* Set outputs *)
stRefTime.dwSec := TIME_TO_DWORD(tonMeassureTime.PT) / 1000;

stRefTime.dwDeciSec := TIME_TO_DWORD(tonMeassureTime.PT) / 100;

stRefTime.dwCentiSec := TIME_TO_DWORD(tonMeassureTime.PT) / 10;

stRefTime.dwMiliSec := TIME_TO_DWORD(tonMeassureTime.PT) / 1;

IF bTimeStarted
THEN
	stActTime.dwSec := stTime.dwSec + TIME_TO_DWORD(tonMeassureTime.ET) / 1000;
	stRestTime.dwSec := TIME_TO_DWORD(tonMeassureTime.PT) / 1000 - stActTime.dwSec;
	
	stActTime.dwDeciSec := stTime.dwDeciSec + TIME_TO_DWORD(tonMeassureTime.ET) / 100;
	stRestTime.dwDeciSec := TIME_TO_DWORD(tonMeassureTime.PT) / 100 - stActTime.dwDeciSec;
	
	stActTime.dwCentiSec := stTime.dwCentiSec + TIME_TO_DWORD(tonMeassureTime.ET) / 10;
	stRestTime.dwCentiSec := TIME_TO_DWORD(tonMeassureTime.PT) / 10 - stActTime.dwCentiSec;

	stActTime.dwMiliSec := stTime.dwMiliSec + TIME_TO_DWORD(tonMeassureTime.ET) / 1;
	stRestTime.dwMiliSec := TIME_TO_DWORD(tonMeassureTime.PT) / 1 - stActTime.dwMiliSec;
END_IF;

IF tonMeassureTime.Q                                		(* Maximum time reached *)
THEN
	MEMSET(ADR(stTime), 0, SIZEOF(stTime));
	bTimeStarted := FALSE;                          		(* Time measure stoped *)
END_IF;

END_FUNCTION_BLOCK

// ---- POUs/Tc2 Objects/Measurements/RTC/FB_RTC.TcPOU
FUNCTION_BLOCK FB_RTC
VAR_INPUT
END_VAR
VAR_OUTPUT
	(* Variables *)
	bTimeValid							:BOOL;
	dtRTC        							:DT;
	dtRTCEX      							:DT;
	stDateTime							:ST_DateTime;
END_VAR
VAR
	(* Enummerations *)

	(* Variables *)
	bFirstTime							:BOOL;	
	bBusy								:BOOL;
	bError								:BOOL;
	udnErrorNo							:UDINT;			

	bValidRTC      						:BOOL;	
	bValidRTCEX    						:BOOL;

	actSysTimeDate						:TIMESTRUCT;				(* Structure SysTimeDate *)
	
	
	(* References *)

	(* Interfaces *)

	(* Instances *)

   	fbGetLocalTime  					:NT_GetTime;
	tonSyncTimer       					:TON;
	ftSyncTrigger     					:F_TRIG;

	rtFirstTime						:R_TRIG;

	fbRTC           						:RTC;
	fbRTCEX        						:RTC_EX;

	(* Information given by the RTC *)
	wYear								:WORD;
	wMonth								:WORD;
	wDay								:WORD;
	wHour								:WORD;
	wMinute								:WORD;
	wSecond							:WORD;
	wMilliseconds						:WORD;

END_VAR

IF NOT bFirstTime
THEN
	bFirstTime := TRUE;
	
END_IF


(* Get RTC *)
rtFirstTime(CLK := bFirstTime);

(* Time synchronization *)
tonSyncTimer(
	IN := NOT tonSyncTimer.Q,
	PT := T#100MS,
);

(* This function provides the time (seconds) which has passed since 01.01.1970 00:00:00 (RTC). *)
fbGetLocalTime(
	NETID := '',
	START := tonSyncTimer.Q
			 OR rtFirstTime.Q,
	TMOUT := T#5S,
	BUSY => bBusy,
	ERR => bError,
	ERRID => udnErrorNo
);

actSysTimeDate := fbGetLocalTime.TIMESTR;

(*This function converts the time given into format SysTimeDate.*)
ftSyncTrigger(CLK := bBusy AND NOT bError);

fbRTC(
	EN := ftSyncTrigger.Q, 
	PDT := SYSTEMTIME_TO_DT(actSysTimeDate), 
	Q => bValidRTC, 
	CDT => dtRTC 
);

fbRTCEX(
	EN := ftSyncTrigger.Q,
	PDT := SYSTEMTIME_TO_DT(actSysTimeDate),
	PMSEK := actSysTimeDate.wMilliseconds,
	Q => bValidRTCEX, 
	CDT => dtRTCEX 
);

(*The structure SysTimeDate contains detailed information on the system time, 
split up into a readable format, e.g.:*)

wYear := actSysTimeDate.wYear;
wMonth := actSysTimeDate.wMonth;
wDay := actSysTimeDate.wDay;
wHour := actSysTimeDate.wHour;
wMinute := actSysTimeDate.wMinute;
wSecond := actSysTimeDate.wSecond;
wMilliseconds := actSysTimeDate.wMilliseconds;

stDateTime.dtDateTime := dtRTC;
stDateTime.dtDateTimeEx := dtRTCEX;

stDateTime.sDate := CONCAT(WORD_TO_STRING(wYear),
		 CONCAT(SEL(LEN(WORD_TO_STRING(wMonth))=1 ,WORD_TO_STRING(wMonth),CONCAT('0',WORD_TO_STRING(wMonth))),
				SEL(LEN(WORD_TO_STRING(wDay))=1 ,WORD_TO_STRING(wDay),CONCAT('0',WORD_TO_STRING(wDay)))));

stDateTime.sTime := CONCAT(SEL(LEN(WORD_TO_STRING(wHour))=1 ,WORD_TO_STRING(wHour),CONCAT('0',WORD_TO_STRING(wHour))),
		 CONCAT(SEL(LEN(WORD_TO_STRING(wMinute))=1 ,WORD_TO_STRING(wMinute),CONCAT('0',WORD_TO_STRING(wMinute))),
				SEL(LEN(WORD_TO_STRING(wSecond))=1 ,WORD_TO_STRING(wSecond),CONCAT('0',WORD_TO_STRING(wSecond)))));

stDateTime.sTimeEx := CONCAT(stDateTime.sTime, SEL(LEN(WORD_TO_STRING(wMilliseconds))=1 , SEL(LEN(WORD_TO_STRING(wMilliseconds))=2 , WORD_TO_STRING(wMilliseconds), CONCAT('0',WORD_TO_STRING(wMilliseconds))), CONCAT('00',WORD_TO_STRING(wMilliseconds))));
				
stDateTime.sDateTime := CONCAT(stDateTime.sDate,CONCAT('_', stDateTime.sTime));

stDateTime.sDateTimeEx := CONCAT(stDateTime.sDate,CONCAT('_', stDateTime.sTimeEx));

END_FUNCTION_BLOCK

// ---- POUs/Tc2 Objects/Traceability/FB_Traceability.TcPOU
FUNCTION_BLOCK FB_Traceability
(*

This function block is used to traceability of data.

Constructor: 		Patryk Panylo
Company:		E. Riexinger GmbH
Date:			02.09.2016
Version:			1.00

Date:			Revision:		Who:				Comment
21.02.2018		0.01			PPA						Additional logger for samples

*)
VAR_INPUT
	(* Input variables / Eingang Variablen *)
	bEnable						:BOOL;					(* Enable FB *)
	bExecute					:BOOL;					(* Execute operation *)
	stTraceability					:ST_Traceability;
END_VAR
VAR_OUTPUT
	(* Output variables / Ausgang Variablen *)
	bBusy						:BOOL;					(* Program busy *)
	bDone						:BOOL;					(* Program done *)
	bError						:BOOL;					(* Program error *)
	udnErrNo					:UDINT;					(* Error number *)
END_VAR
VAR
	(* Enummerations *)

	(* Variables *)
	sDateTimeCache				:STRING;
	arsDataRecord				:ARRAY[0..udnTraceSampleMax] OF STRING(udnTraceStringLengthMax);
	udnDataRecordCnt			:UDINT;

	udnIdxData					:UDINT;
	udnIdxSample				:UDINT;
	enStep						:INT;

	bFirstTime					:BOOL;					(* First PLC cycle *)

	(* References *)

	(* Interfaces *)

	(* Instances *)
	fbTraceability					:FB_FileHandler;				(* Traceability *)
	rtExecute						:R_TRIG;
END_VAR
VAR CONSTANT
	sEndLine					:STRING := '$N'; 							(* End line sign for lines *)
END_VAR

IF NOT bEnable				(* Enable FB *)
THEN
	bFirstTime := FALSE;		(* First PLC cycle *)
	bBusy := FALSE;			(* Program busy *)
	bDone := FALSE;			(* Program done *)
	bError := FALSE;			(* Program error *)
	udnErrNo := 0;				(* Error number *)
	RETURN;
END_IF

IF NOT bFirstTime
THEN

	bFirstTime := TRUE;
END_IF

rtExecute(CLK := bExecute);

IF rtExecute.Q
    AND NOT fbTraceability.bBusy
THEN
	sDateTimeCache := stTraceability.sDateTime;

	FOR udnIdxSample := 0 TO udnTraceSampleMax
	DO

		IF udnIdxSample = 0
		THEN
			arsDataRecord[udnIdxSample] := CONCAT('No', sTraceColSep);

			FOR udnIdxData := 1 TO udnTraceDataMax
			DO
				IF LEN(stTraceability.arstData[1,udnIdxData].sName) <> 0
				     AND LEN(stTraceability.arstData[1,udnIdxData].sValue) <> 0
				THEN
					arsDataRecord[udnIdxSample] := CONCAT(arsDataRecord[udnIdxSample],
											  			   CONCAT(stTraceability.arstData[1,udnIdxData].sName,
													  			    CONCAT(' ',
															 			     CONCAT(stTraceability.arstData[1,udnIdxData].sUnit, sTraceColSep)
													 					     )
											  					    )
														 );

				END_IF

				IF udnIdxData = udnTraceDataMax
				    AND LEN(arsDataRecord[udnIdxSample]) <> 0
				THEN
					arsDataRecord[udnIdxSample] := REPLACE(arsDataRecord[udnIdxSample], sEndLine, 1, LEN(arsDataRecord[udnIdxSample]));
				END_IF
			END_FOR

		ELSE

			arsDataRecord[udnIdxSample] := CONCAT(UDINT_TO_STRING(udnIdxSample), sTraceColSep);
	
			FOR udnIdxData := 1 TO udnTraceDataMax
			DO
				IF LEN(stTraceability.arstData[udnIdxSample,udnIdxData].sName) <> 0
				     AND LEN(stTraceability.arstData[udnIdxSample,udnIdxData].sValue) <> 0
				THEN
					arsDataRecord[udnIdxSample] := CONCAT(arsDataRecord[udnIdxSample],
												CONCAT(stTraceability.arstData[udnIdxSample,udnIdxData].sValue, sTraceColSep)
											);
		
				END_IF
		
				IF udnIdxData = udnTraceDataMax
				    AND LEN(arsDataRecord[udnIdxSample]) <> 0
				THEN
					arsDataRecord[udnIdxSample] := REPLACE(arsDataRecord[udnIdxSample], sEndLine, 1, LEN(arsDataRecord[udnIdxSample]));
				END_IF
			END_FOR

		END_IF

	END_FOR
END_IF

CASE enStep
OF

	0:
		IF rtExecute.Q
		THEN
			udnDataRecordCnt := 0;
			fbTraceability.sWriteRecord := arsDataRecord[udnDataRecordCnt];

			enStep := 1;
		END_IF

	1:
		fbTraceability.bExecute := TRUE;

		IF fbTraceability.bBusy
		     AND NOT fbTraceability.bError
		THEN

			enStep := 2;
		ELSIF fbTraceability.bError
		THEN
			fbTraceability.bExecute := FALSE;

			enStep := 0;
		END_IF
	2:
		IF fbTraceability.bDone
		     AND NOT fbTraceability.bError
		THEN
			fbTraceability.bExecute := FALSE;

			enStep := 3;

		ELSIF fbTraceability.bError
		THEN
			fbTraceability.bExecute := FALSE;

			enStep := 0;
		END_IF

	3:	IF NOT fbTraceability.bBusy
		     AND NOT fbTraceability.bDone
		     AND NOT fbTraceability.bError
		THEN
			fbTraceability.bExecute := FALSE;

			udnDataRecordCnt := udnDataRecordCnt +1;
			IF udnDataRecordCnt < udnTraceSampleMax
			THEN
				fbTraceability.sWriteRecord := arsDataRecord[udnDataRecordCnt];

				enStep := 1;
			ELSE
				enStep := 0;
			END_IF

		ELSIF fbTraceability.bError
		THEN
			fbTraceability.bExecute := FALSE;

			enStep := 0;
		END_IF

END_CASE

fbTraceability(
	bEnable := TRUE,
	sFilePath := stTraceability.stSettings.sPath,
	sFileName := CONCAT(sDateTimeCache, (*CONCAT('_', stTraceability.stSettings.sFileName)*)''),
	sFileSuffix := stTraceability.stSettings.sFileExtension,
	dwOpenMode := FOPEN_MODEAPPEND (* OR  FOPEN_MODETEXT*),
	tTimeout := t#2s,
	bBusy => bBusy,
	bDone => bDone,
	bError => bError,
	udnErrNo => udnErrNo);

END_FUNCTION_BLOCK

// ---- POUs/Tc2 Objects/File/FB_FileHandler.TcPOU
FUNCTION_BLOCK FB_FileHandler
(*

This function block is used to read and write binary datas in/from file.

Constructor: 		Patryk Panylo
Company:		E. Riexinger GmbH
Date:			10.06.2013
Version:			1.00

Date:			Revision:		Who:				Comment
dd.mm.yyyy		x.xx			Initials			comment

*)

VAR_INPUT
	bEnable						:BOOL;					(* Enable FB *)
	bExecute					:BOOL;					(* Execute operation *)
	sFilePath					:STRING;				(* File path *)
	sFileName					:STRING;				(* File name *)
	sFileSuffix					:STRING := 'dat';			(* Suffix of file *)
	dwOpenMode				:DWORD;				(*
															FOPEN_MODEREAD (16#0001)	"r": Opens for reading. If the file does not exist or cannot be found, the call fails.
															FOPEN_MODEWRITE (16#0002) "w": Opens an empty file for writing. If the given file exists, its contents are destroyed.
															FOPEN_MODEAPPEND (16#0004) "a": Opens for writing at the end of the file (appending) without removing the EOF marker before writing new data to the file; creates the file first if it doesn’t exist.
															FOPEN_MODEREAD OR FOPEN_MODEPLUS (16#0008) "r+": Opens for reading and writing. The file must exist.
															FOPEN_MODEWRITE OR FOPEN_MODEPLUS (16#0008) "w+": Opens an empty file for both reading and writing. If the given file exists, its contents are destroyed.
															FOPEN_MODEAPPEND OR FOPEN_MODEPLUS (16#0008)	 "a+": Opens for reading and appending; the appending operation includes the removal of the EOF marker before new data is written to the file and the EOF marker is restored after writing is complete; creates the file first if it doesn’t exist.
															When a file is opened with the "a" or "a+" access type, all write operations occur at the end of the file. The file pointer can be repositioned using FB_FileSeek, but is always moved back to the end of the file before any write operation is carried out. Thus, existing data cannot be overwritten.
															
															FOPEN_MODEBINARY (16#0010) "b": Open in binary (untranslated) mode.
															FOPEN_MODETEXT (16#0020) "t": Open in text (translated) mode.
														*)
	sWriteRecord					:T_MaxString;				(* Record to write *)
	tTimeout						:TIME := t#1s;				(* States the time before the function is cancelled *)
END_VAR
VAR_OUTPUT
	sReadRecord				:T_MaxString;				(* Record to read *)
	bBusy						:BOOL;					(* Program busy *)
	bDone						:BOOL;					(* Program done *)
	bError						:BOOL;					(* Program error *)
	udnErrNo					:UDINT;					(* Error number *)
END_VAR
VAR_IN_OUT

END_VAR
VAR
	(* Enummerations *)
	enStep						: (eWaitExecute := 0, eChkFileName,  eChkBufLen, eCreateDir, eChkCreateDir, eFileOpen, eChkFileOpen, eFileWrite, eChkFileWrite, eFileRead, eChkFileRead, eFileClose, eChkFileClose, eDone, eError, eNotExecute);			(* Sequence state for open, read/write and close the file *)

	(* Variables *)
	bFirstTime					:BOOL;					(* First PLC cycle *)

	dwModeCache				:DWORD;				(* Contains the mode in which the file is to be opened *)
	sWriteRecordCache			:T_MaxString;				(* Record to write *)
	sPathName					:STRING;				(* Contains the path and filename for the file to be opened *)
	hFileHandle					:UINT;					(* File handle *)

	unWriteCounter				:UINT;
	unReadCounter				:UINT;

	(* Instances *)
	fbCreateDir					:FB_CreateDir;			(* File open *)
	fbFileOpen					:FB_FileOpen;			(* File open *)
	fbFileClose					:FB_FileClose;			(* File close *)
	fbFileRead					:FB_FileRead;			(* File read *)
	fbFileWrite					:FB_FileWrite;				(* File write *)

END_VAR

IF NOT bEnable				(* Enable FB *)
THEN
	bFirstTime := FALSE;		(* First PLC cycle *)
	bBusy := FALSE;			(* Program busy *)
	bDone := FALSE;			(* Program done *)
	bError := FALSE;			(* Program error *)
	udnErrNo := 0;				(* Error number *)
	RETURN;
END_IF

IF NOT bFirstTime
THEN
	enStep := eWaitExecute;

	bFirstTime := TRUE;
END_IF


(* Sequence state for open, read/write and close the file *)
CASE enStep
OF

	eWaitExecute:
		IF bExecute
		THEN
			fbFileOpen.bExecute := FALSE;			(* File open *)
			fbFileClose.bExecute := FALSE;			(* File close *)
			fbFileRead.bExecute := FALSE;			(* File read *)
			fbFileWrite.bExecute := FALSE;			(* File write *)

			bDone := FALSE;
			bError := FALSE;
			udnErrNo := 0;

			sWriteRecordCache := sWriteRecord;

			IF dwOpenMode <> 0
			THEN
				dwModeCache := dwOpenMode;

				enStep := eChkFileName;			(* Next step *)

			ELSE
				RETURN;
			END_IF

			bBusy := TRUE;

		END_IF

	(* Check file name and path *)
	eChkFileName:

		sPathName := CONCAT(
						sFilePath, CONCAT(
									sFileName, CONCAT(
												'.', sFileSuffix)));

		IF sFilePath <> ''
		     AND sFileName <> ''
		     AND sFileSuffix <> ''
		THEN
			enStep := eChkBufLen;			(* Next step *)

		ELSE
			udnErrNo := eChkFileName;

			enStep := eError;				(* Next step *)

		END_IF


	(* Check buffer lenght *)
	eChkBufLen:
		IF LEN(sWriteRecordCache) = 0
		THEN
			enStep := eDone;				(* Next step *)
	
		ELSE
			(*enStep := eCreateDir;			(* Next step *)*)
			enStep := eFileOpen;			(* Next step *)
		END_IF

	(* Create direction *)
	eCreateDir:
		fbCreateDir.bExecute := TRUE;

		enStep := eChkCreateDir;				(* Next step *)

	eChkCreateDir:
		IF NOT fbCreateDir.bBusy
		THEN
			IF NOT fbCreateDir.bError
			THEN
				fbCreateDir.bExecute := FALSE;

				enStep := eFileOpen;				(* Next step *)
			ELSE
				fbCreateDir.bExecute := FALSE;

				IF  fbCreateDir.nErrId = 16#70C 	(* 0x70C Folder is allready existing or invalid sPathName or ePath parameter.*)
				THEN
					enStep := eFileOpen;				(* Next step *)
				ELSE
					enStep := eError;					(* Next step *)
				END_IF
			END_IF
		END_IF

	(* Open the file *)
	eFileOpen:
		IF LEN(sWriteRecordCache) > 254
		THEN
			sWriteRecordCache := DELETE(
								sWriteRecordCache,
								LEN(sWriteRecordCache) + 1 - 254, 254
							    );
		END_IF

		fbFileOpen.bExecute := TRUE;

		enStep := eChkFileOpen;				(* Next step *)

	(* Check open the file *)
	eChkFileOpen:
		IF NOT fbFileOpen.bBusy
		THEN
			IF NOT fbFileOpen.bError
			THEN
				fbFileOpen.bExecute := FALSE;
				hFileHandle := fbFileOpen.hFile;

				(* Choose write or read datas *)
				IF fbFileOpen.nMode = FOPEN_MODEWRITE
				THEN
				
					enStep := eFileWrite;			(* Next step *)

				ELSIF fbFileOpen.nMode = FOPEN_MODEAPPEND
				THEN
	
					enStep := eFileWrite;			(* Next step *)

				ELSIF fbFileOpen.nMode = FOPEN_MODEREAD
				THEN
					enStep := eFileRead;			(* Next step *)
				
				ELSE
					enStep := eFileClose;			(* Next step *)

				END_IF

			ELSE
				fbFileOpen.bExecute := FALSE;
				udnErrNo := fbFileOpen.nErrId;
	
				enStep := eError;					(* Next step *)
				
			END_IF
		END_IF

	(* Write the file *)
	eFileWrite:
		fbFileWrite.bExecute := TRUE;

		enStep := eChkFileWrite;				(* Next step *)

	(* Check write the file *)
	eChkFileWrite:
		IF NOT fbFileWrite.bBusy
		THEN
			IF (fbFileWrite.cbWrite >= INT_TO_UDINT(LEN(sWriteRecordCache)))
			    AND NOT fbFileWrite.bError
			THEN
				fbFileWrite.bExecute := FALSE;
				unWriteCounter := unWriteCounter + 1;

				enStep := eFileClose;				(* Next step *)

			ELSIF  fbFileWrite.bError
			THEN
				fbFileWrite.bExecute := FALSE;
				udnErrNo := fbFileWrite.nErrId;

				enStep := eError;					(* Next step *)
				
			END_IF
		END_IF

	(* Read the file *)
	eFileRead:
		fbFileRead.bExecute := TRUE;

		enStep := eChkFileRead;				(* Next step *)

	(* Check read the file *)
	eChkFileRead:
		IF NOT fbFileRead.bBusy
		THEN
			IF (fbFileRead.cbRead >= INT_TO_UDINT(LEN(sReadRecord)))
			     AND NOT fbFileRead.bError
			THEN
				fbFileRead.bExecute := FALSE;
				unReadCounter := unReadCounter + 1;
	
				enStep := eFileClose;				(* Next step *)

			ELSIF  fbFileRead.bError
			THEN
				fbFileRead.bExecute := FALSE;
				udnErrNo := fbFileRead.nErrId;
	
				enStep := eError;					(* Next step *)
				
			END_IF
		END_IF

	(* Close the file *)
	eFileClose:
		fbFileClose.bExecute := TRUE;

		enStep := eChkFileClose;				(* Next step *)

	(* Check close the file *)
	eChkFileClose:
		IF NOT fbFileClose.bBusy
		THEN
			IF NOT fbFileClose.bError
			THEN
				fbFileClose.bExecute := FALSE;
				enStep := eDone;					(* Next step *)

				IF bError
				THEN
					enStep := eError;				(* Next step *)
				END_IF

			ELSE
				fbFileClose.bExecute := FALSE;
				udnErrNo := fbFileClose.nErrId;
	
				enStep := eError;					(* Next step *)
				
			END_IF
		END_IF

	eDone:
		bBusy := FALSE;
		bDone := TRUE;
		bError := FALSE;
		udnErrNo := 0;

		enStep := eNotExecute;					(* Next step *)

	eError:
		IF NOT bError
		     AND hFileHandle <> 0
		THEN
			bDone := FALSE;
			bError := TRUE;

			enStep := eFileClose;					(* Next step *)

		ELSE
			bBusy := FALSE;
			bDone := FALSE;
			bError := TRUE;
	
			enStep := eNotExecute;					(* Next step *)
		END_IF

	eNotExecute:
		IF NOT bExecute
		THEN
			bBusy := FALSE;
			bDone := FALSE;
			bError := FALSE;
			udnErrNo := 0;

			enStep := eWaitExecute;			(* Next step *)

		END_IF

END_CASE

fbCreateDir(
	sNetId:= '',
	sPathName:= sFilePath,
	ePath:= PATH_GENERIC,
	tTimeout:= tTimeout);
fbFileOpen(
	sNetId := '',
	sPathName := sPathName,
	nMode := dwModeCache,
	ePath := PATH_GENERIC,
	tTimeout := tTimeout);
fbFileClose(
	sNetId := '',
	hFile := hFileHandle,
	tTimeout := tTimeout );
fbFileWrite(
	sNetId := '',
	hFile := hFileHandle,
	pWriteBuff := ADR(sWriteRecordCache),
	cbWriteLen := INT_TO_UDINT(LEN(sWriteRecordCache)),
	tTimeout := tTimeout);
fbFileRead(
	sNetId := '',
	hFile := hFileHandle,
	pReadBuff := ADR(sReadRecord),
	cbReadLen := INT_TO_UDINT(LEN(sReadRecord)),
	tTimeout := tTimeout);

END_FUNCTION_BLOCK

// ---- POUs/Machine/Group_0000 - General/Gr00Control/Gr00Periphery/FB_Gr00Periphery.TcPOU
FUNCTION_BLOCK FB_Gr00Periphery
(*

The function block used to control periphery.

Constructor: 		Patryk Panylo
Company:		E. Riexinger GmbH
Date:			24.10.2015
Version:			1.00

Date:			Revision:		Who:				Comment
dd.mm.yyyy		x.xx			Initials			comment

*)
VAR_INPUT
	(* Input variables / Eingang Variablen *)
	bEnable						:BOOL;						(* Axis present *)
END_VAR
VAR_OUTPUT
	(* Output variables / Ausgang Variablen *)

END_VAR
VAR_IN_OUT
	(* Input Output variables / Ausgang Variablen *)
	Periphery					:FB_PERIPHERY_REF;			(* Interface of periphery *)
END_VAR
VAR
	(* Enummerations *)

	(* Variables *)

	(* References *)

	(* Interfaces *)

	(* Instances *)

END_VAR

IF NOT bEnable								(* Signal FB enable *)
THEN

	RETURN;
END_IF

A_PeripheryLink();

ACTION A_PeripheryLink:

;
END_ACTION

END_FUNCTION_BLOCK

// ---- POUs/Tc2 Objects/ExternalHardware/Periphery/FB_PERIPHERY_REF.TcPOU
FUNCTION_BLOCK FB_PERIPHERY_REF
VAR_INPUT

END_VAR
VAR_OUTPUT

END_VAR
VAR_IN_OUT

END_VAR
VAR

END_VAR

;

END_FUNCTION_BLOCK

// ---- POUs/Tc2 Objects/Signals/Handling/FB_SignalHandlingDelay.TcPOU
FUNCTION_BLOCK FB_SignalHandlingDelay
VAR_INPUT
	(* Input variables / Eingang Variablen *)
	bEnable					:BOOL;						(* Enable FB signal *)
	bIn						:BOOL;						(* Input signal *)
	tDelay					:TIME := t#0s;					(* Delay *)
END_VAR
VAR_OUTPUT
	(* Output variables / Ausgang Variablen *)
	bOut					:BOOL;						(* Delayed signal *)
END_VAR
VAR
	(* Enummerations *)

	(* Variables *)
	bFirstTime				:BOOL;						(* First cycle *)

	(* References *)

	(* Interfaces *)

	(* Instances *)
	tonDelay					:TON;						(* Timer to delay *)
END_VAR

IF NOT bEnable
THEN
	tonDelay(IN := FALSE,
	          	PT := tDelay);
	bOut := bIn;
    RETURN;
END_IF;

tonDelay(				(* Dealy input signal *)
	IN := bIn,
	PT := tDelay
);

bOut := tonDelay.Q;		(* Set output *)

END_FUNCTION_BLOCK

// ---- POUs/Machine/Group_0100 - Production/Gr01MachineMode/Gr01Home/Gr01Home.TcPOU
PROGRAM Gr01Home
VAR_INPUT
	(* Input variables / Eingang Variablen *)
	bEnable					:BOOL;						(* Enable Gr05Home *)
	bExecute				:BOOL;						(* Home execute *)

	(* Instances *)
	fbInit						:FB_Gr01HomeInit;
	fbProcedure				:FB_Gr01HomeProcedure;

	fbAxisSawBow			:FB_Gr01HomeAxisSawBow;
	fbAxisAngle				:FB_Gr01HomeAngle;
	fbSawband				:FB_Gr01HomeSawband;

END_VAR
VAR
	(* Enummerations *)

	(* Variables *)

	(* References *)

	(* Interfaces *)

	(* Instances *)
	rtExecute					:R_TRIG;

	fbAlarm					:FB_Gr01HomeAlarm;

END_VAR
VAR CONSTANT
	nFatalErrorMaxIdx				:INT := 0;						(* Maximal index of  using alarms *)
	nErrorMaxIdx					:INT := 1;						(* Maximal index of  using alarms *)
	nWarningMaxIdx				:INT := 0;						(* Maximal index of  using alarms *)
	nMessageMaxIdx				:INT := 0;						(* Maximal index of  using alarms *)
	nHintMaxIdx					:INT := 0;						(* Maximal index of  using alarms *)

	dnFatalErrorBaseIdentNo		:DINT := 13000;				(* Fatal error identification number *)
	dnErrorBaseIdentNo			:DINT := 13100;				(* Error identification number *)
	dnWarningBaseIdentNo		:DINT := 13200;				(* Warning identification number *)
	dnMessageBaseIdentNo		:DINT := 13300;				(* Message identification number *)
	dnHintBaseIdentNo			:DINT := 13400;				(* Hint identification number *)
END_VAR

IF NOT bEnable
THEN
	RETURN;
END_IF;

(* Check home execute *)
bExecute := etgGr00MachineState = ET_MachineState_eHomeRefExe
		      OR etgGr00MachineState = ET_MachineState_eHomeExe;

rtExecute(CLK := bExecute);

IF rtExecute.Q
THEN
	fbInit.bFirstTime := FALSE;
	A_Init();
END_IF;

A_Procedure();
A_Functions();
A_Alarm();

ACTION A_Alarm:

(* Collect and execute input alarms *)
fbAlarm.stAlarmIn.arbError[0].bActive := fbAxisSawBow.bErrorByReference;
fbAlarm.stAlarmIn.arbError[0].dnCode := dnErrorBaseIdentNo + 0;

fbAlarm.stAlarmIn.arbError[1].bActive := fbAxisAngle.bErrorByReference;
fbAlarm.stAlarmIn.arbError[1].dnCode := dnErrorBaseIdentNo + 1;

fbAlarm(
	etMachineMode := etgGr00MachineMode,
	etMachineState := etgGr00MachineState,
	bNoEStop := bgGr00NoEmergencyStop,
	bConfirmAlarm := bgGr00ConfirmAlarm,
	dtDateTime := stgGr00DateTime.dtDateTime,
	nFatalErrorMaxIdx := nFatalErrorMaxIdx,
	nErrorMaxIdx := nErrorMaxIdx,
	nWarningMaxIdx := nWarningMaxIdx,
	nMessageMaxIdx := nMessageMaxIdx,
	nHintMaxIdx := nHintMaxIdx,
	bMoveInterrupted := bgGr01MoveInterrupted,
	bHomeCompleted := bgGr01HomeCompleted,
	stAlarmOut => stgGr01Alarm.stHome
);
END_ACTION

ACTION A_Functions:

fbAxisSawBow(
	bEnable := etgGr00MachineMode = ET_MachineMode_eHome,
	bReleaseNextStep := etgGr00MachineState = ET_MachineState_eHomeRefExe
		      	     		      OR etgGr00MachineState = ET_MachineState_eHomeExe,
	pfbAxis := ADR(Gr01Control.fbAxisSawBow)
);

fbAxisAngle(
	bEnable := etgGr00MachineMode = ET_MachineMode_eHome,
	bReleaseNextStep := etgGr00MachineState = ET_MachineState_eHomeRefExe
		      	     		      OR etgGr00MachineState = ET_MachineState_eHomeExe,
	pfbAxis := ADR(Gr01Control.fbAxisAngle)
);

fbSawband(
	bEnable := etgGr00MachineMode = ET_MachineMode_eHome,
	bReleaseNextStep := etgGr00MachineState = ET_MachineState_eHomeRefExe
		      	     		      OR etgGr00MachineState = ET_MachineState_eHomeExe,
	pfbAxis := ADR(Gr01Control.fbSawband)
);
END_ACTION

ACTION A_Init:

(* Initializing variables *)
fbInit();
END_ACTION

ACTION A_Procedure:

(* Execute home procedure *)
fbProcedure(
	bEnable := etgGr00MachineMode = ET_MachineMode_eHome,
	bExecute := rtExecute.Q,
	bReleaseNextStep := etgGr00MachineState = ET_MachineState_eHomeRefExe
		      	     		      OR etgGr00MachineState = ET_MachineState_eHomeExe
);
END_ACTION

END_PROGRAM

// ---- POUs/Machine/Group_0100 - Production/Gr01Control/Gr01Control.TcPOU
PROGRAM Gr01Control
VAR_INPUT
	(* Input variables / Eingang Variablen *)
	bEnable						:BOOL;						(* Enable Gr01Control *)

	(* Instances *)
	fbAxisSawBow				:FB_Gr01SawBow;
	fbAxisAngle					:FB_Gr01Angle;

	fbSawband			 		:FB_Gr01Sawband;

END_VAR
VAR
	(* Enummerations *)

	(* Variables *)
	bAllAxisCtrlEnabled				:BOOL;						(* All axis have controller enabled *)
	bAllAxisStandStill				:BOOL;						(* All axis stand still *)
	bAllAxisNotMoving				:BOOL;						(* All axis not moving *)
	bAllAxisReferenced				:BOOL;						(* All axis referenced *)
	
	BandDistance_m					:LREAL;
	rMachineSawbandSpeed_mmin		:LREAL;

	(* References *)

	(* Interfaces *)

	(* Instances *)
	fbAlarm						:FB_Gr01Alarm;
	fbSafety					:FB_Gr01Safety;
	fbSignals					:FB_Gr01Signals;
	fbUtility					:FB_Gr01Utility;
	rtBtnStart					:R_TRIG;
	
	SawbandVelo					:FB_PosVeloEnc;
	fbLowPassFilter				:FB_LowPassFilter;
	tonSawBandVeloErr			:TON;
	tonSawBandInVelo			:TON;
	TimerVelo					:TON;

END_VAR
VAR CONSTANT
	nFatalErrorMaxIdx			:INT := 0;						(* Maximal index of  using alarms *)
	nErrorMaxIdx				:INT := 19;					(* Maximal index of  using alarms *)
	nWarningMaxIdx				:INT := 0;						(* Maximal index of  using alarms *)
	nMessageMaxIdx				:INT := 1;						(* Maximal index of  using alarms *)
	nHintMaxIdx					:INT := 0;						(* Maximal index of  using alarms *)

	dnFatalErrorBaseIdentNo		:DINT := 11000;				(* Fatal error identification number *)
	dnErrorBaseIdentNo			:DINT := 11100;				(* Error identification number *)
	dnWarningBaseIdentNo		:DINT := 11200;				(* Warning identification number *)
	dnMessageBaseIdentNo		:DINT := 11300;				(* Message identification number *)
	dnHintBaseIdentNo			:DINT := 11400;				(* Hint identification number *)
END_VAR

IF NOT bEnable
THEN
	RETURN;
END_IF;

A_Utility();
A_Safety();
A_Axis();
A_Sawband();
A_Signals();
A_Alarm();

ACTION A_Alarm:

(* Collect and execute input alarms *)
fbAlarm.stAlarmIn.arbError[0].bActive := NOT binGr01LightCurtainOK
                                                		      AND (Gr01Home.fbProcedure.bBusy
                                                      				OR Gr01Auto.fbProcedure.bBusy);
fbAlarm.stAlarmIn.arbError[0].dnCode := dnErrorBaseIdentNo + 0;

fbAlarm.stAlarmIn.arbError[1].bActive := NOT binGr01SawbandRelease
								    AND bgGr00ModeAutomatic
								    AND bgGr00MachineRunning;
fbAlarm.stAlarmIn.arbError[1].dnCode := dnErrorBaseIdentNo + 1;

fbAlarm.stAlarmIn.arbError[2].bActive := FALSE;
fbAlarm.stAlarmIn.arbError[2].dnCode := dnErrorBaseIdentNo + 2;

fbAlarm.stAlarmIn.arbError[3].bActive := FALSE;
fbAlarm.stAlarmIn.arbError[3].dnCode := dnErrorBaseIdentNo + 3;

fbAlarm.stAlarmIn.arbError[4].bActive := fbAxisSawBow.bErrorTerminal;
fbAlarm.stAlarmIn.arbError[4].dnCode := dnErrorBaseIdentNo + 4;

fbAlarm.stAlarmIn.arbError[5].bActive := fbAxisSawBow.fbController.bErrorInit;
fbAlarm.stAlarmIn.arbError[5].dnCode := dnErrorBaseIdentNo + 5;

fbAlarm.stAlarmIn.arbError[6].bActive := fbAxisSawBow.bErrorCtrlEnabled;
fbAlarm.stAlarmIn.arbError[6].dnCode := dnErrorBaseIdentNo + 6;

fbAlarm.stAlarmIn.arbError[7].bActive := fbAxisSawBow.fbController.bError OR fbAxisSawBow.fbMoveManual.bError OR fbAxisSawBow.fbMoveAuto.bError;
fbAlarm.stAlarmIn.arbError[7].dnCode := dnErrorBaseIdentNo + 7;

fbAlarm.stAlarmIn.arbError[8].bActive := fbAxisAngle.bErrorTerminal;
fbAlarm.stAlarmIn.arbError[8].dnCode := dnErrorBaseIdentNo + 8;

fbAlarm.stAlarmIn.arbError[9].bActive := fbAxisAngle.fbController.bErrorInit;
fbAlarm.stAlarmIn.arbError[9].dnCode := dnErrorBaseIdentNo + 9;

fbAlarm.stAlarmIn.arbError[10].bActive := fbAxisAngle.bErrorCtrlEnabled;
fbAlarm.stAlarmIn.arbError[10].dnCode := dnErrorBaseIdentNo + 10;

fbAlarm.stAlarmIn.arbError[11].bActive := fbAxisAngle.fbController.bError OR fbAxisAngle.fbMoveManual.bError OR fbAxisAngle.fbMoveAuto.bError;
fbAlarm.stAlarmIn.arbError[11].dnCode := dnErrorBaseIdentNo + 11;

fbAlarm.stAlarmIn.arbError[12].bActive := fbSawband.bErrorTerminal;
fbAlarm.stAlarmIn.arbError[12].dnCode := dnErrorBaseIdentNo + 12;

fbAlarm.stAlarmIn.arbError[13].bActive := fbSawband.fbController.bErrorInit;
fbAlarm.stAlarmIn.arbError[13].dnCode := dnErrorBaseIdentNo + 13;

fbAlarm.stAlarmIn.arbError[14].bActive := fbSawband.bErrorCtrlEnabled;
fbAlarm.stAlarmIn.arbError[14].dnCode := dnErrorBaseIdentNo + 14;

fbAlarm.stAlarmIn.arbError[15].bActive := fbSawband.fbController.bError OR fbSawband.fbMoveManual.bError OR fbSawband.fbMoveAuto.bError;
fbAlarm.stAlarmIn.arbError[15].dnCode := dnErrorBaseIdentNo + 15;

fbAlarm.stAlarmIn.arbError[16].bActive := FALSE;
fbAlarm.stAlarmIn.arbError[16].dnCode := dnErrorBaseIdentNo + 16;

fbAlarm.stAlarmIn.arbError[17].bActive := GVL_Gr0100.bgGr01SawbandVeloError_1;
fbAlarm.stAlarmIn.arbError[17].dnCode := dnErrorBaseIdentNo + 17;

fbAlarm.stAlarmIn.arbError[18].bActive := GVL_Gr0100.bgGr01SawbandVeloError_2;
fbAlarm.stAlarmIn.arbError[18].dnCode := dnErrorBaseIdentNo + 18;

fbAlarm.stAlarmIn.arbError[19].bActive := (* bgGr00MachineRunning
							AND fbSawband.bCtrlEnabled
							AND fbSawband.bSpeedReached
							AND *) NOT fbSafety.bPipeNotInCrashArea;  (* 20260219 ES/KG *)

fbAlarm.stAlarmIn.arbError[19].dnCode := dnErrorBaseIdentNo + 19;

fbAlarm.stAlarmIn.arbWarning[0].bActive := fbSawband.bErrorVacuumCleanerNOK;
fbAlarm.stAlarmIn.arbWarning[0].dnCode := dnWarningBaseIdentNo + 0;

fbAlarm.stAlarmIn.arbMessage[0].bActive := NOT binGr01LightCurtainOK
							      AND NOT fbAlarm.stAlarmIn.arbError[0].bActive
							      AND NOT fbAlarm.stAlarmOut.arbError[0].bActive;
fbAlarm.stAlarmIn.arbMessage[0].dnCode := dnMessageBaseIdentNo + 0;

fbAlarm.stAlarmIn.arbMessage[1].bActive := NOT binGr01SawbandRelease;
fbAlarm.stAlarmIn.arbMessage[1].dnCode := dnMessageBaseIdentNo + 1;

(* Execute utility *)
fbAlarm(
	etMachineMode := etgGr00MachineMode,
	etMachineState := etgGr00MachineState,
	bNoEStop := bgGr00NoEmergencyStop,
	bConfirmAlarm := bgGr00ConfirmAlarm,
	dtDateTime := stgGr00DateTime.dtDateTime,
	nFatalErrorMaxIdx := nFatalErrorMaxIdx,
	nErrorMaxIdx := nErrorMaxIdx,
	nWarningMaxIdx := nWarningMaxIdx,
	nMessageMaxIdx := nMessageMaxIdx,
	nHintMaxIdx := nHintMaxIdx,
	bMoveInterrupted := bgGr01MoveInterrupted,
	bHomeCompleted := bgGr01HomeCompleted,
	stAlarmOut => stgGr01Alarm.stControl
);
END_ACTION

ACTION A_Axis:

(* Enable axis saw bow *)
stgGr01HMI.stHMITOPLC.lrAxisSawBowNoRefVelo := 10;

fbAxisSawBow(
	bEnable						:= TRUE,
	etMachineMode				:= etgGr00MachineMode,
	etMachineState				:= etgGr00MachineState,
	bMachineStandstill			:= bgGr00MachineStandstill,
	bNoEStop					:= bgGr00NoEmergencyStop,
	bPowerSupplyOn				:= bgGr00PowerSupplyOk,
	bSafetyOK					:= bgGr01LightCurtainOK
								   AND bgGr00AllDoorsClosedLocked,
	bCtrlInterrupt				:= FALSE,
	bMoveRelease				:= TRUE,
	bPlusRelease				:= TRUE,
	bMinusRelease				:= TRUE,
	bSignalReference			:= NOT binGr01AxisSawBowLimitMax,
	bSignalHWLimitMax			:= NOT binGr01AxisSawBowLimitMax,
	bSignalHWLimitMin			:= NOT binGr01AxisSawBowLimitMin,
	lrSoftLimitMax				:= stgGr01HMI.stHMITOPLC.lrAxisSawBowSoftLimitMax,
	lrSoftLimitMin				:= stgGr01HMI.stHMITOPLC.lrAxisSawBowSoftLimitMin,
	bConfirmAlarm				:= bgGr00ConfirmAlarm,
	bTipPlus					:= stgGr01HMI.stHMITOPLC.bBtnAxisSawBowPlus,
	bTipMinus					:= stgGr01HMI.stHMITOPLC.bBtnAxisSawBowMinus,
	lrManualVelocity			:= stgGr01HMI.stHMITOPLC.lrAxisSawBowManualVelo,
	lrNoRefVelocity				:= stgGr01HMI.stHMITOPLC.lrAxisSawBowNoRefVelo,
	bVelocityLimitEn			:= FALSE,
	lrAcceleration				:= 100.0,
	lrDeceleration				:= 100.0,
	lrJerk						:= 100.0,
	lrOverride					:= fbUtility.rActOverride,
	lrExtOverride				:= 0.0,
	dnRatioNumerator			:= 1,
	udnRatioDenominator			:= 1,
	bEngineTorqueLimitEn		:= FALSE,
	lrEngineTorque				:= 200.0,
	tControllerOff				:= tgGr01ControllerOff,
	bWithAbsoluteEncoder		:= FALSE,
	lrOriginShiftPos			:= stgGr01HMI.stHMITOPLC.lrAxisSawBowOriginShiftPos,
	bVeloForceCtrlEn			:= FALSE,
	tAdsTimeOut					:= DEFAULT_ADS_TIMEOUT,
	bHomeCompleted				:= bgGr01HomeCompleted,
	Drive						:= GVL_Gr01Interface.igGr01DriveSawBow,
	Axis						:= GVL_Gr01Interface.igGr01AxisSawBow,
	MasterAxis					:= GVL_Gr00Interface.iAxisDummy,
	
	lrActPosition				=> stgGr01HMI.stPLCTOHMI.lrAxisSawBowActPos,
	lrActVelocity				=> stgGr01HMI.stPLCTOHMI.lrAxisSawBowActVelo,
	lrActForce					=> stgGr01HMI.stPLCTOHMI.lrAxisSawBowActForce
);

(* Enable Axis angle *)
stgGr01HMI.stHMITOPLC.lrAxisAngleNoRefVelo := 10;



fbAxisAngle(
	bEnable						:= TRUE,

	etMachineMode				:= etgGr00MachineMode,
	etMachineState				:= etgGr00MachineState,
	bMachineStandstill			:= bgGr00MachineStandstill,
	bNoEStop					:= bgGr00NoEmergencyStop,
	bPowerSupplyOn				:= bgGr00PowerSupplyOk,
	bSafetyOK					:= bgGr01LightCurtainOK
								   AND bgGr00AllDoorsClosedLocked,
	bCtrlInterrupt				:= FALSE,
	bMoveRelease				:= TRUE,
	bMoveInterrupt				:= FALSE,
	bPlusRelease				:= TRUE,
	bMinusRelease				:= TRUE,	(*stgGr00HMI.stHMITOPLC.bSafetyInterlockOff*)
	bHWSignalLimitMax			:= NOT binGr01AxisAngleLimitMax,
	bHWSignalLimitMin			:= NOT binGr01AxisAngleLimitMin,
	lrSoftLimitMax				:= stgGr01HMI.stHMITOPLC.lrAxisAngleSoftLimitMax,
	lrSoftLimitMin				:= stgGr01HMI.stHMITOPLC.lrAxisAngleSoftLimitMin,
	bConfirmAlarm				:= bgGr00ConfirmAlarm,
	bTipPlus					:= stgGr01HMI.stHMITOPLC.bBtnAxisAnglePlus,
	bTipMinus					:= stgGr01HMI.stHMITOPLC.bBtnAxisAngleMinus,
	lrManualVelocity			:= stgGr01HMI.stHMITOPLC.lrAxisAngleManualVelo,
	lrVelocityNoRef				:= stgGr01HMI.stHMITOPLC.lrAxisAngleNoRefVelo,
	bVelocityLimitEn			:= FALSE,
	lrAcceleration				:= 100.0,
	lrDeceleration				:= 100.0,
	lrJerk						:= 100.0,
	lrOverride					:= fbUtility.rActOverride,
	bEngineTorqueLimitEn		:= FALSE,
	lrEngineTorque				:= 200.0,
	tControllerOff				:= tgGr01ControllerOff,
	lrScalingNum				:= lrgGr01AxisAnglePath,
	udnScalingDenom				:= udngGr01AxisAngleInc,
	bWithAbsoluteEncoder		:= TRUE,
	udnIncEnc					:= udninGr01IncAxisAngle,
	lrOriginShift				:= stgGr01HMI.stHMITOPLC.lrAxisAngleOriginShiftPos,
	lrTaskCycle					:= lrgActCycleTime,
	tAdsTimeOut					:= DEFAULT_ADS_TIMEOUT,
	bHomeCompleted				:= bgGr01HomeCompleted,
	Drive						:= GVL_Gr01Interface.igGr01DriveSawAngle,
	Axis						:= GVL_Gr01Interface.igGr01AxisSawAngle,
	MasterAxis					:= GVL_Gr00Interface.iAxisDummy,
	
	lrActPosition				=> stgGr01HMI.stPLCTOHMI.lrAxisAngleActPos,
	lrActVelocity				=> stgGr01HMI.stPLCTOHMI.lrAxisAngleActVelo
);
END_ACTION

ACTION A_Safety:

(* Execute safety *)
fbSafety(
	bLightCurtain := binGr01LightCurtainOK,
	bConfirmLightCurtain := (bgGr00ConfirmAlarm
			                            OR etgGr00MachineMode = ET_MachineMode_eManual
			                            OR etgGr00MachineMode = ET_MachineMode_eHome
			                            OR etgGr00MachineMode = ET_MachineMode_eAutomatic
			                            OR stgGr00HMI.stHMITOPLC.bSafetyInterlockOff)
					         AND NOT stgGr01Alarm.stControl.arbError[0].bActive,
	tLightCurtainDelay := tgGr01LightCurtainDelay,
	bLightCurtainOK => bgGr01LightCurtainOK,
	bConfirmedLightCurtain => boutGr01ConfLightCurtain,
	bNotInCrashArea => bgGr01NotInCrashArea
);

bgGr01SafetyActive := fbAxisSawBow.bSafetyLock
				        OR fbAxisAngle.bSafetyLock;
END_ACTION

ACTION A_Sawband:

fbSawband(
	bEnable						:= TRUE,
	bOccupied					:= FALSE,
	etMachineMode				:= etgGr00MachineMode,
	etMachineState				:= etgGr00MachineState,
	bMachineStandstill			:= bgGr00MachineStandstill,
	bNoEStop					:= bgGr00NoEmergencyStop,
	bPowerSupplyOn				:= bgGr00PowerSupplyOk,	//fbStoeberPS6A34.bOn, // Keine Eingänge vorhanden
	bSafetyOK					:= bgGr01LightCurtainOK								   AND bgGr00AllDoorsClosedLocked,
	bSafetyDriveEnabled			:= TRUE,
	bCtrlInterrupt				:= FALSE,
	bMoveRelease				:= TRUE,
	bPlusRelease				:= TRUE,
	bMinusRelease				:= FALSE,
	bSignalReference			:= FALSE,
	bSignalHWLimitMax			:= FALSE,
	bSignalHWLimitMin			:= FALSE,
	lrSoftLimitMax				:= 0,
	lrSoftLimitMin				:= 0,
	etHomingMode				:= MC_DefaultHoming,
	bConfirmAlarm				:= bgGr00ConfirmAlarm,
	bTipPlus					:= stgGr01HMI.stHMITOPLC.bBtnSawbandPlus,
	bTipMinus					:= False,
	lrTipDistance				:= 0,
	lrManualVelocity			:= stgGr01HMI.stHMITOPLC.rSawbandManualSpeed / 3.28084,
	lrAutoVelocity				:= stgGr01HMI.stHMITOPLC.rSawbandAutoSpeed / 3.28084,
	lrNoRefVelocity				:= 30,
	bVelocityLimitEn			:= FALSE,
	lrAcceleration				:= 5000,
	lrDeceleration				:= 5000,
	lrJerk						:= 30000,
	lrOverride					:= 100.0,
	bExtOverrideEn				:= FALSE,
	dnRatioNumerator			:= 1,
	udnRatioDenominator			:= 1,
	bEngineTorqueLimitEn		:= FALSE,
	lrEngineTorque				:= 400,
	bPosLagMonitoringEn			:= FALSE,
	tControllerOff				:= tgGr01ControllerOff,
	bWithAbsoluteEncoder		:= FALSE,
	bVeloForceCtrlEn			:= FALSE,
	tAdsTimeOut					:= DEFAULT_ADS_TIMEOUT,
	bHomeCompleted				:= bgGr01HomeCompleted,
	Drive						:= GVL_Gr01Interface.igGr01DriveSawBand,
	Axis						:= GVL_Gr01Interface.igGr01AxisSawBand,
	MasterAxis					:= GVL_Gr00Interface.iAxisDummy,

	lrActVelocity				=> GVL_Gr01HMI.stgGr01HMI.stPLCTOHMI.lrSawbandActSpeed,
	bSawbandAirOn 				=> boutGr01SawbandAirOn
);

rMachineSawbandSpeed_mmin := stgGr01HMI.stHMITOPLC.rSawbandAutoSpeed / 3.28084;

////////////// Sawband Velo Scaling

SawbandVelo(
	bEnable				:= TRUE , 
	dwEncCurrentValue	:= GVL_GR01IO.udninGr01CounterSawbandSpeed, 
	udnScalingDenom		:= uiImpulsDiscAmount , 	
	lrScalingNum		:= rRaddurchmesser_mm*PI, 	
	tCycleTime			:= GVL_Gr00Init.tPLC_TaskCycleTime_ms, 					
	lrCurrentPos		=> , 
	lrCurrentVelo		=> ,			(* [mm/ms] same as [m/s]*)
);
	
BandDistance_m := SawbandVelo.lrCurrentPos / 1000;
GVL_Gr01Init.lrgGr01SawingSpeed := SawbandVelo.lrCurrentVelo * 60;		(* [m/min] *)

	fbLowPassFilter(
	bEnable			:= TRUE , 
	lrIn			:= GVL_Gr01Init.lrgGr01SawingSpeed, 
	lrKp			:= 1, 
	tT1				:= T#600MS , 
	tCycletime		:= GVL_Gr00Init.tPLC_TaskCycleTime_ms, 
	lrOut			=> GVL_Gr01Init.lrgGr01SawingSpeed

);
//////////////
GVL_Gr01HMI.stgGr01HMI.stHMITOPLC.rSawbandAutoSpeed := GVL_Gr01Init.lrgGr01SawingSpeed;
	
	
////////////// Sawband Velo Error -> never reaches target speed
tonSawBandInVelo(
					IN:= NOT GVL_GR0100.bgGr01SawbandVeloError_1 AND (ABS(GVL_Gr01Interface.igGr01AxisSawBand.NcToPlc.ActVelo) - ABS(GVL_Gr01Interface.igGr01AxisSawBand.NcToPlc.SetVelo)< 100),
					PT := T#3S);
					
GVL_GR0100.bgGr01SawbandInSpeed := GVL_Gr01Init.lrgGr01SawingSpeed > (rMachineSawbandSpeed_mmin * 0.8 * fbSawband.lrOverride/100)
							AND (tonSawBandInVelo.Q OR GVL_Gr01HMI.stgGr01HMI.stHMITOPLC.bBtnSawbandPlus);
							
TimerVelo(
	IN:= NOT GVL_GR0100.bgGr01SawbandInSpeed AND NOT GVL_GR0100.bgGr01SawbandVeloError_1 AND GVL_Gr0000.bgGr00NoEmergencyStop, 
	PT:=T#10S
		); 
		
GVL_GR0100.bgGr01SawbandVeloError_1 := TimerVelo.Q; 


//Sawband velocity error -> lost target speed
tonSawBandVeloErr(
					IN:=ABS(GVL_Gr01Interface.igGr01AxisSawBand.NcToPlc.ActVelo) < ABS(GVL_Gr01Interface.igGr01AxisSawBand.NcToPlc.SetVelo *0.8),
					PT := T#500MS);

GVL_GR0100.bgGr01SawbandVeloError_2 := tonSawBandInVelo.Q;



(* Old FB)
(* Enable sawband *)
fbSawband(
	bEnable := TRUE,
	lrScalingNum := lrgGr01SawbandDistance,
	udnScalingDenom := udngGr01SawbandInc,
	etMachineMode := etgGr00MachineMode,
	etMachineState := etgGr00MachineState,
	bNoEStop := bgGr00NoEmergencyStop,
	bPowerSupplyOn := bgGr00PowerSupplyOk,
	bSafetyOK := bgGr01LightCurtainOK
			        AND bgGr00AllDoorsClosedLocked,
	bAirPressureOK := bgGr00AirPressureOK,
	bMachineStandstill := bgGr00MachineStandstill,
	bCtrlInterrupt := FALSE,
	bMoveRelease := TRUE,
	bMoveInterrupt := FALSE,
	bTipPlus := stgGr01HMI.stHMITOPLC.bBtnSawbandPlus,
	bTipMinus := FALSE(*stgGr01HMI.stHMITOPLC.bBtnSawbandMinus*),
	bPlusRelease := TRUE,
	bMinusRelease := TRUE,
	bHandSawbandAirOn := stgGr01HMI.stHMITOPLC.bBtnSawbandAirOn,
	bHandVacuumCleanerOn := stgGr01HMI.stHMITOPLC.bBtnVacuumCleanerOn,
	bExtOverrideEn := FALSE,
	lrManualSpeed := stgGr01HMI.stHMITOPLC.rSawbandManualSpeed / 3.28084,
	lrAutoSpeed := stgGr01HMI.stHMITOPLC.rSawbandAutoSpeed  / 3.28084,
	bSpeedLimitEn := TRUE,
	lrSpeedMin := 0, (* m/min *)
	lrSpeedMax := 400, (* m/min  SY 650*)
	lrAcceleration := 100.0,
	lrDeceleration := 100.0,
	lrJerk := 100.0,
	bEngineTorqueLimitEn := FALSE,
	lrEngineTorque := 200.0,
	bSawbandMotorNOK := binGr01SawbandMotorNOK,
	bSawbandBroken := NOT binGr01SawbandNoBroken,
	bVacuumCleanerMotorNOK := binGr01VacuumCleanerMotorNOK,
	udnIncEnc := udninGr01CounterSawbandSpeed,
	lrTaskCycle := lrgActCycleTime,
	bConfirmAlarm := bgGr00ConfirmAlarm,
	tSawbandAirOffDelay := tgGr01SawbandAirOffDelay,
	tVacuumCleanerOffDelay := tgGr01VacuumCleanerOffDelay,
	tSawbandReadyDelay := tgGr01SawbandReadyDelay,
	tSpeedNoConstant := tgGr01SpeedNoConstant,
	tControllerOff := tgGr01ControllerOff,
	tAdsTimeOut := DEFAULT_ADS_TIMEOUT,
	bHomeCompleted := bgGr01HomeCompleted,
	Drive := igGr01DriveSawband,
	Axis := igGr01AxisSawband,
	lrActSpeed => stgGr01HMI.stPLCTOHMI.lrSawbandActSpeed,
	bSawbandAirOn => boutGr01SawbandAirOn,
	bVacuumCleanerOn => boutGr01VacuumCleanerOn
);
*)
END_ACTION

ACTION A_Signals:

(* Execute signals *)
fbSignals(
	etMachineMode := etgGr00MachineMode,
	etMachineState := etgGr00MachineState,
	bMachineRunning := bgGr00MachineRunning,
	bExecutedProcess := fbUtility.arbExeProcess[1]
					      OR fbUtility.arbExeProcess[2]
					      OR fbUtility.arbExeProcess[3],
	stBlinker := stgGr00Blinker,
	bBulbBtnStart => boutGr01BulbBtnStart,
	bBulbBtnStop => boutGr01BulbBtnStop,
);

(* Detect all axis controller enabled *)
bAllAxisCtrlEnabled := F_ChkAllAxisEnabled(
	bEnable := TRUE,
	bEnabledAxis1 := Gr01Control.fbAxisSawBow.bCtrlEnabled,
	bEnabledAxis2 := Gr01Control.fbAxisAngle.bCtrlEnabled,
	bEnabledAxis3 := TRUE,
	bEnabledAxis4 := TRUE,
	bEnabledAxis5 := TRUE,
	bEnabledAxis6 := TRUE,
	bEnabledAxis7 := TRUE,
	bEnabledAxis8 := TRUE,
	bEnabledAxis9 := TRUE,
	bEnabledAxis10 := TRUE
);

(* Detect all axis stand still *)
bAllAxisStandStill := F_ChkAllAxisStandStill(
	bEnable := TRUE,
	bAxis1StandStill := Gr01Control.fbAxisSawBow.bStandStill, 		// igGr01AxisSawBow.stAxisStatus.bStandStill,
	bAxis2StandStill := Gr01Control.fbAxisAngle.bStandStill,		// igGr01AxisAngle.stAxisStatus.bStandStill,
	bAxis3StandStill := TRUE,
	bAxis4StandStill := TRUE,
	bAxis5StandStill := TRUE,
	bAxis6StandStill := TRUE,
	bAxis7StandStill := TRUE,
	bAxis8StandStill := TRUE,
	bAxis9StandStill := TRUE,
	bAxis10StandStill := TRUE,
);

(* Detect all axis not moving *)
bAllAxisNotMoving := F_ChkAllAxisNotMoving(
	bEnable := TRUE,
	bAxis1NotMoving := Gr01Control.fbAxisSawBow.bNotMoving, 		
	bAxis2NotMoving := Gr01Control.fbAxisAngle.bNotMoving,
	bAxis3NotMoving := TRUE,
	bAxis4NotMoving := TRUE,
	bAxis5NotMoving := TRUE,
	bAxis6NotMoving := TRUE,
	bAxis7NotMoving := TRUE,
	bAxis8NotMoving := TRUE,
	bAxis9NotMoving := TRUE,
	bAxis10NotMoving := TRUE
);

(* Detect all axis referenced *)
bAllAxisReferenced := F_ChkAllAxisReferenced(
	bEnable := TRUE,
	bReferencedAxis1 := Gr01Control.fbAxisSawBow.bReferenced,
	bReferencedAxis2 := Gr01Control.fbAxisAngle.bReferenced,
	bReferencedAxis3 := TRUE,
	bReferencedAxis4 := TRUE,
	bReferencedAxis5 := TRUE,
	bReferencedAxis6 := TRUE,
	bReferencedAxis7 := TRUE,
	bReferencedAxis8 := TRUE,
	bReferencedAxis9 := TRUE,
	bReferencedAxis10 := TRUE
);
END_ACTION

ACTION A_Utility:

(* Execute utility *)

(* Start program *)
rtBtnStart(CLK := binGr00PushBtnStart OR stgGr00HMI.stHMITOPLC.bBtnStart);

fbUtility.arbStartProcess[1] := rtBtnStart.Q
						 AND etgGr00MachineState = ET_MachineState_eAutoExe;
fbUtility.arbStopProcess[1] := etgGr00MachineState <> ET_MachineState_eAutoExe;
fbUtility.arbSteppingProcess[1] := stgGr01HMI.stHMITOPLC.bBtnSteppingProcess;
arbgGr01StartProcess[1] := fbUtility.arbExeProcess[1];

fbUtility(
	etMachineMode := etgGr00MachineMode,
	etMachineState := etgGr00MachineState,
	bAutoCompleted := bgGr00AutoCompleted
					  AND bgGr01AutoCompleted
					  AND bgGr02AutoCompleted
					  AND bgGr05AutoCompleted
					  AND bgGr00MachineStandstill
					  AND etgGr00MachineState <> ET_MachineState_eAutoExe,
	bHomeCompleted := bgGr01HomeCompleted,
	bExeCounter := bgGr01AutoCompleted,
	bLaserOnOff := stgGr01HMI.stHMITOPLC.bBtnLaserOn,
	bStartTime := Gr01Control.fbUtility.arbStartProcess[1]
				OR Gr01Control.fbUtility.arbStartProcess[2]
				OR Gr01Control.fbUtility.arbStopProcess[3],
	bStopTime := bgGr01AutoCompleted
				OR fbUtility.arbStopProcess[1]
				OR fbUtility.arbStopProcess[2]
				OR fbUtility.arbStopProcess[3],
	bLifetimeOn := NOT fbSawband.bNotMoving,
	bResetLifetimeAll := FALSE,
	bResetLifetime := stgGr01HMI.stHMITOPLC.bResetLifetime,
	sLifetimeFilePath := sgGr01LifetimeFilePath,
	sLifetimeFileName := sgGr01LifetimeFileName,
	bPipeIdentify := NOT binGr01PipeNoIdentify,
	rGlobalOverride := rgGr00Override,
	rLocalOverride := stgGr01HMI.stHMITOPLC.rOverride,
	lrLifetimeAll => stgGr01HMI.stPLCTOHMI.lrLifetime,
	lrLifetimeAfterReset => stgGr01HMI.stPLCTOHMI.lrLifetimeAfterReset,
	lrLifetimeAfterTrunOn => stgGr01HMI.stPLCTOHMI.lrLifetimeAfterTurnOn,
	udnCounterTotal := stgGr01HMI.stPLCTOHMI.udnCounterTotal,
	bLaserOn => boutGr01LaserOn,
	bPipePresent => bgGr01PipePresent
);
END_ACTION

END_PROGRAM

// ---- POUs/Machine/Group_0100 - Production/Gr01Control/Gr01Units/FB_Gr01SawBow.TcPOU
FUNCTION_BLOCK FB_Gr01SawBow
(*

The function block used to control axis welding.

Constructor: 		Patryk Panylo
Company:			E. Riexinger GmbH
Date:				28.04.2015
Version:			1.00

Date:			Revision:		Who:				Comment
dd.mm.yyyy		x.xx			Initials			comment

*)
VAR_INPUT
	(* Input variables / Eingang Variablen *)

	(* --- Axis / Achse --- *)
	bEnable						:BOOL;						(* Axis present *)
	bOccupied					:BOOL;						(* Axis occupied *)

	(* --- Machine state / Maschinenzustand --- *)
	etMachineMode				:ET_MachineMode;			(* Machine mode *)
	etMachineState				:ET_MachineState;			(* Machine state *)
	bMachineStandstill			:BOOL;						(* Machine standstill *)

	(* --- Safety & releases / Sicherheit & Freigaben --- *)
	bNoEStop					:BOOL;						(* No ermergency Stop / Keine Notaus *)
	bPowerSupplyOn				:BOOL;						(* Power supply on / Leitung eingeschaltet *)
	bSafetyOK					:BOOL;						(* Safety ok / Sicherheit i.o *)
	bSafetyDriveEnabled			:BOOL;						(* Safety drive enable *)
	bCtrlInterrupt				:BOOL;						(* Control interrupt *)
	bMoveRelease				:BOOL;						(* Move release *)
	bPlusRelease				:BOOL;						(* Plus move release *)
	bMinusRelease				:BOOL;						(* Minus move release *)

	(* --- Limits & signals / Endlagen & Signale --- *)
	bSignalReference			:BOOL;						(* Reference signal *)
	bSignalHWLimitMax			:BOOL;						(* Position Hard limit switch maximum *)
	bSignalHWLimitMin			:BOOL;						(* Position Hard limit switch minimum *)
	lrSoftLimitMax				:LREAL;						(* Position limit switch maximum *)
	lrSoftLimitMin				:LREAL;						(* Position limit switch minimum *)

	(* --- Commands / Befehle --- *)
	bExeReset					:BOOL;						(* Execute auto reset *)
	bExeCtrlEnable				:BOOL;						(* Controller enable *)
	bExeSetPos					:BOOL;						(* Execute set position *)
	bExeHome					:BOOL;						(* Execute home *)
	etHomingMode				:MC_HomingMode;				(* HomingMode determines in which way the calibration is carried out. *)
	bExeMoveAbs					:BOOL;						(* Execute move absolut *)
	bExeMoveRel					:BOOL;						(* Execute move relative *)
	bExeMoveAdd					:BOOL;						(* Execute move additive *)
	bExeMoveSuper				:BOOL;						(* Execute move superimposed *)
	bExeMoveVelo				:BOOL;						(* Execute move velo *)
	bExeGearIn					:BOOL;						(* Execute gear in *)
	bExeGearOut					:BOOL;						(* Execute gear out *)
	bExeStop					:BOOL;						(* Execute move stop *)
	bConfirmAlarm				:BOOL;						(* Confirm alarm *)

	(* --- Manual mode / Handbetrieb --- *)
	bTipPlus					:BOOL;						(* Manual tip in plus direction *)
	bTipMinus					:BOOL;						(* Manual tip in minus direction *)
	lrTipDistance				:LREAL;						(* Relative distance for movements *)
	lrManualVelocity			:LREAL;						(* Value of velocity in manual motion [mm/s] *)

	(* --- Motion parameters / Bewegungsparameter --- *)
	lrTargetPosition			:LREAL;						(* Absolute target position *)
	lrTargetPositionOffset		:LREAL;						(* Absolute target position offset *)
	lrAutoVelocity				:LREAL;						(* Value of velocity in auto motion [mm/s] *)
	lrNoRefVelocity				:LREAL;						(* Velocity if has no reference [mm/s] *)
	bVelocityLimitEn			:BOOL;						(* Enable velocity limit *)
	lrVelocityMin				:LREAL;						(* Velocity minimum [%] *)
	lrVelocityMax				:LREAL;						(* Velocity maximum [%] *)
	lrAcceleration				:LREAL;						(* Value of the acceleration (always positive) *)
	lrDeceleration				:LREAL;						(* Value of deceleration (always positive) *)
	lrJerk						:LREAL;						(* Value of jerk (always positive) *)

	(* --- Override --- *)
	lrOverride					:LREAL;						(* Override *)
	bExtOverrideEn				:BOOL;						(* External override enable *)
	lrExtOverride				:LREAL;						(* External override *)

	(* --- Gearing / Getriebe --- *)
	dnRatioNumerator			:DINT;						(* Gear ratio numerator. Alternatively, the gear ratio can be specified in the numerator as a floating comma value, if the denominator is 1. *)
	udnRatioDenominator			:UDINT;						(* Gear ratio denominator *)

	(* --- Drive / Antrieb --- *)
	snModesOfOperation			:SINT;						(* Modes of drive operation *)
	bEngineTorqueLimitEn		:BOOL;						(* Enable engine torque limit *)
	lrEngineTorque				:LREAL;						(* Engine torque [%] *)
	bPosLagMonitoringEn			:BOOL;						(* Enable position lag monitoring *)
	tControllerOff				:TIME := T#60S;				(* Time to switch controller off *)

	(* --- Encoder / Geber --- *)
	bWithAbsoluteEncoder		:BOOL;						(* Encoder is an absolute one / Absolutwertgeber *)
	lrOriginShiftPos			:LREAL;						(* Origin shift position *)

	(* --- Force control / Kraftregelung --- *)
	unForceMeasureType			:UINT;						(* Type of force measure system. 1: Simple mA,  2: EL3351 3: EL3356 *)
	bVeloForceCtrlEn			:BOOL;						(* Enable velocity  force controller *)
	lrVeloForceCtrlKp			:LREAL;						(* Velocity - force controller proportional band Kp *)
	lrVeloForceCtrlTi			:LREAL;						(* Velocity - force controller integral Ti *)
	lrVeloForceCtrlMin			:LREAL;						(* Velocity - force controller minimum  *)
	lrVeloForceCtrlMax			:LREAL;						(* Velocity - force controller maxmimum  *)
	lrVeloForcePreCtrlVelo		:LREAL;						(* Feedforward velocity precontrol wieghting =  0..1 *)
	lrTargetForce				:LREAL;						(* Absolute target force [N] *)
	lrForceCurrent				:LREAL;						(* Current force [mA] *)
	rForceOffset				:REAL;						(* Force offset [N] *)
	lrMaintenanceOverflowForce	:LREAL;						(* Maintenance overflow force [N] *)
	lrManualOverflowForce		:LREAL;						(* Maximal force in manual mode [N] *)
	lrAutoOverflowForce			:LREAL;						(* Maximal force in automatic mode [N] *)
	lrForceMinmA				:LREAL;						(* Force min [mA] 16#0000 = 4 [mA] *)
	lrForceMaxmA				:LREAL;						(* Force max [mA] 16#7FFF = 20 [mA] *)
	lrForceMinN					:LREAL;						(* Force min [N] *)
	lrForceMaxN					:LREAL;						(* Force max [N] *)

	(* --- Temperature & cooling / Temperatur & Kühlung --- *)
	lrActTemp					:LREAL;						(* Current temperatur *)
	lrTempLimitMax				:LREAL;						(* Temperatur limit maximum*)
	lrTempLimitMin				:LREAL;						(* Temperatur limit minimum*)
	bCoolingActive				:BOOL;						(* Cooling on *)

	(* --- System --- *)
	tAdsTimeOut					:TIME := T#2S;				(* Timout for ads commands *)
END_VAR
VAR_OUTPUT
	(* Output variables / Ausgang Variablen *)

	(* --- Status --- *)
	bCtrlEnabled				:BOOL;						(* Controller enabled *)
	bNotMoving					:BOOL;						(* Axis not moving *)
	bStandStill					:BOOL;						(* Added by Dustin for 633_Hilton) Axis stands stil*)
	bReferenced					:BOOL;						(* Axis referenced *)
	bCoupled					:BOOL;						(* Axis coupled *)

	(* --- Actual values / Istwerte --- *)
	lrActPosition				:LREAL;						(* Actual position [mm] *)
	lrActAbsPosition			:LREAL;						(* Actual absolut position [mm] *)
	lrActVelocity				:LREAL;						(* Actual velocity [mm/s] *)
	lrActForce					:LREAL;						(* Actual force [N] *)
	lrVeloMax					:LREAL;						(* Velocity limit maximum *)
	lrAccMax					:LREAL;						(* Acceleration limit maximum *)
	lrDecMax					:LREAL;						(* Deceleration limit maximum *)
	lrJerkMax					:LREAL;						(* Jerk limit maximum *)

	(* --- Limits / Endlagen --- *)
	bHardLimitMaxExceeded		:BOOL;						(* Position limit switch maximum is exceeded *)
	bHardLimitMinExceeded		:BOOL;						(* Position limit switch minimum is exceeded *)
	bSoftLimitMaxExceeded		:BOOL;						(* Position limit switch maximum is exceeded *)
	bSoftLimitMinExceeded		:BOOL;						(* Position limit switch minimum is exceeded *)

	(* --- Peripherals / Peripherie --- *)
	bCoolingOn					:BOOL;						(* Cooling *)

	(* --- Safety / Sicherheit --- *)
	bSafetyLock					:BOOL;						(* Safety lock*)
	bSafetyDriveEnable			:BOOL;						(* Safety drive enable *)

	(* --- Errors / Fehler --- *)
	bErrorTerminal				:BOOL;						(* Error Axis terminal *)
	bErrorDrive					:BOOL;						(* Error drive *)
	bErrorCtrlEnabled			:BOOL;						(* Error Axis controller enabled *)
	bErrorForceOverflow			:BOOL;						(* Error force overflow *)
	bErrPosLimitOverflow		:BOOL;						(* Error position limit overflow *)
END_VAR
VAR_IN_OUT
	(* Input Output variables / Ausgang Variablen *)
	bHomeCompleted				:BOOL;						(* Home completed *)
	Drive						:ST_STOEBERSI6SC6CIA402_REF; (* The ST_STOEBERSI6SC6CIA402_REF data type  is an interface between the PLC and the DRIVE and contains axis information *)
	Axis						:AXIS_REF;					(* The AXIS_REF data type  is an interface between the PLC and the NC and contains axis information *)
	MasterAxis					:AXIS_REF;					(* The AXIS_REF data type  is an interface between the PLC and the NC and contains axis information *)
END_VAR
VAR
	(* Enummerations *)

	(* Variables *)
	sAdsAddr					:STRING(23);					(* AmsNetId of the EtherCAT master device.*)
	unSlaveAddr					:UINT;						(* Address of the slave device.*)

	nTorqueLimitMax				:INT := 100;					(* The torque limit (absolute value). Value range in %: -200 ... 200 ... 200 *)

	lrVeloLimitMax				:LREAL;
	lrVeloLimitMin				:LREAL;

	sTerminalStatus				:STRING;
	
	bSetCoeParaToDefault		:BOOL;
	bReadCoePara				:BOOL;
	bWriteCoePara				:BOOL;
	stCoeWrite					:ST_EL3356CoeInfo;
	stCoeRead					:ST_EL3356CoeInfo;
	
	lrCacheWeightTara			:LREAL;
	
	(* References *)

	(* Interfaces *)

	(* Instances *)
	fbTerminalDiagnosis			:FB_TerminalDiagnosis;
	rtMachineStandstill			:R_TRIG;
	tonAxisEnabled				:TON;

